CheckInitialization := FSetupValid
    AND FEqualResult.IsInitialized
    AND FNotEqualResult.IsInitialized
    AND FCaptureIntegrity.IsInitialized
    AND FFindingDetails.IsInitialized;
IF NOT CheckInitialization THEN
    EventPublisher.PublishEvent(Event := CreateFrameworkEvent(Name := Name,
        ResourceName := '',
        State := State,
        Severity := E_EventSeverity.Error,
        Message := 'Tolerance selftest setup failed.'));
END_IF;
END_METHOD

{region 'Documentation'}
(*!
<summary>Checks literal results, finding count and isolated finding identities.</summary>
*)
{endregion}
METHOD PRIVATE CheckResults
VAR
    FindingIndex : UINT;
    NotEqualFindingMatches : BOOL;
END_VAR
FEqualResultMatches := FEqualSubject.Result = FExpectedEqualResult;
FNotEqualResultMatches := FNotEqualSubject.Result = FExpectedNotEqualResult;
FCaptureIntegrityMatches := (FCaptureStatus.SequenceId = FExpectedFindings)
    AND (FCaptureStatus.LostEventCount = 0);

FindingIndex := 1;
FFindingDetailsMatch := TRUE;
IF FExpectedEqualFinding <> E_Result.NotEvaluated THEN
    FFindingDetailsMatch := IsFindingValid(Index := FindingIndex,
        ExpectedName := FEqualSubject.Name,
        ExpectedResult := FExpectedEqualFinding);
    FindingIndex := FindingIndex + 1;
END_IF;
IF FExpectedNotEqualFinding <> E_Result.NotEvaluated THEN
    NotEqualFindingMatches := IsFindingValid(Index := FindingIndex,
        ExpectedName := FNotEqualSubject.Name,
        ExpectedResult := FExpectedNotEqualFinding);
    FFindingDetailsMatch := FFindingDetailsMatch AND NotEqualFindingMatches;
END_IF;
END_METHOD

{region 'Documentation'}
(*!
<summary>Configures checking Assertions; subject actions remain in the test script.</summary>
*)
{endregion}
METHOD PROTECTED Configure
VAR
    Initialized : BOOL;
END_VAR
FPreparationStateCount := 0;
FTestStateCount := 1;
FEqualResult.Initialize(Parent := THIS^,
    AssertionName := 'EqualResult');
FNotEqualResult.Initialize(Parent := THIS^,
    AssertionName := 'NotEqualResult');
FCaptureIntegrity.Initialize(Parent := THIS^,
    AssertionName := 'CaptureIntegrity');
FFindingDetails.Initialize(Parent := THIS^,
    AssertionName := 'FindingDetails');
FSetupValid := FCapture.Initialize(Buffer := FEvents,
    FifoControl := FCaptureFifo,
    Status := FCaptureStatus);
FEqualSubject.BindPublisher(Publisher := FCapture);
Initialized := FEqualSubject.Initialize(Parent := THIS^,
    AssertionName := 'EqualSubject');
FSetupValid := FSetupValid AND Initialized;
FNotEqualSubject.BindPublisher(Publisher := FCapture);
Initialized := FNotEqualSubject.Initialize(Parent := THIS^,
    AssertionName := 'NotEqualSubject');
FSetupValid := FSetupValid AND Initialized;
END_METHOD

{region 'Documentation'}
(*!
<summary>Reads one of at most two captured findings; caller supplies index 1 or 2.</summary>
*)
{endregion}
METHOD PRIVATE IsFindingValid : BOOL //! TRUE when the selected captured finding satisfies the scenario metadata and diagnostic checks.
VAR_INPUT
    Index : UINT; //! One-based index in the retained isolated event capture.
    ExpectedName : STRING(GVL_Constants.NameLength); //! Independently authored Assertion name expected in the selected finding.
    ExpectedResult : E_Result; //! Independently authored finding result.
END_VAR
IsFindingValid := (FEvents[Index].SequenceId = UINT_TO_UDINT(Index))
    AND (FEvents[Index].Name = ExpectedName)
    AND (FEvents[Index].OwnerScope = E_OwnerScope.Assertion)
    AND (FEvents[Index].EventType = E_EventType.Result)
    AND (FEvents[Index].State = E_State.Running)
    AND (FEvents[Index].Result = ExpectedResult)
    AND (FEvents[Index].Message <> '');
END_METHOD

{region 'Documentation'}
(*!
<summary>Completes abort without asynchronous resources.</summary>
*)
{endregion}
METHOD PROTECTED ProcessAbort
VAR_INPUT
    Enable : BOOL; //! Phase permission supplied by the owning Test Case; FALSE does not authorize progression, while observation may continue.
END_VAR
IF Enable THEN
    CompleteAbort();
END_IF;
END_METHOD

{region 'Documentation'}
(*!
<summary>Latches checked observations before the next script step may proceed.</summary>
*)
{endregion}
METHOD PROTECTED ProcessAssertions
VAR_INPUT
    Enable : BOOL; //! Phase permission supplied by the owning Test Case; FALSE does not authorize progression, while observation may continue.
END_VAR
VAR
    Evaluate : BOOL;
END_VAR
Evaluate := Enable AND FObservationReady;
FEqualResult(Enable := Evaluate,
    State := State,
    IN := FEqualResultMatches);
FNotEqualResult(Enable := Evaluate,
    State := State,
    IN := FNotEqualResultMatches);
FCaptureIntegrity(Enable := Evaluate,
    State := State,
    IN := FCaptureIntegrityMatches);
FFindingDetails(Enable := Evaluate,
    State := State,
    IN := FFindingDetailsMatch);
IF Evaluate THEN
    FChecked := TRUE;
END_IF;
END_METHOD

{region 'Documentation'}
(*!
<summary>No Preparation phase is required.</summary>
*)
{endregion}
METHOD PROTECTED ProcessPreparations
VAR_INPUT
    // SA0033: Required hook; this test has no Preparation phase.
    {attribute 'analysis' := '-33'}
    Enable : BOOL; //! Phase permission supplied by the owning Test Case; FALSE does not authorize progression, while observation may continue.
END_VAR
END_METHOD

{region 'Documentation'}
(*!
<summary>Restarts the script and resets the checking Assertions.</summary>
*)
{endregion}
METHOD PROTECTED ProcessReset
FRow := EqualValues;
FRowPrepared := FALSE;
FChecked := FALSE;
FObservationReady := FALSE;
FEqualResult.Reset();
FEqualResultMatches := TRUE;
FNotEqualResult.Reset();
FNotEqualResultMatches := TRUE;
FCaptureIntegrity.Reset();
FCaptureIntegrityMatches := TRUE;
FFindingDetails.Reset();
FFindingDetailsMatch := TRUE;
CompleteReset();
END_METHOD

{region 'Documentation'}
(*!
<summary>Advances one bounded script step per active PLC cycle.</summary>
*)
{endregion}
METHOD PROTECTED ProcessTests
VAR_INPUT
    Enable : BOOL; //! Phase permission supplied by the owning Test Case; FALSE does not authorize progression, while observation may continue.
END_VAR
IF NOT Enable THEN
    RETURN;
END_IF;

IF FChecked THEN
    FChecked := FALSE;
    FObservationReady := FALSE;
    IF FRow = LastRow THEN
        CompleteTests();
        RETURN;
    END_IF;
    FRow := FRow + 1;
    FRowPrepared := FALSE;
END_IF;

IF NOT FRowPrepared THEN
    SelectRow();
    FCapture.Reset();
    IF NOT FPreserveResults THEN
        ResetSubjects();
    END_IF;
    CallSubjects(Enable := FALSE);
    FRowPrepared := TRUE;
ELSE
    CallSubjects(Enable := TRUE);
    CheckResults();
    FObservationReady := TRUE;
END_IF;
END_METHOD

{region 'Documentation'}
(*!
<summary>Requests fresh subject results before the next disabled call.</summary>
*)
{endregion}
METHOD PRIVATE ResetSubjects
FEqualSubject.Reset();
FNotEqualSubject.Reset();
END_METHOD

{region 'Documentation'}
(*!
<summary>Selects literal expectations; only named escalation rows retain preceding subject results.</summary>
*)
{endregion}
METHOD PRIVATE SelectRow
FPreserveResults := FALSE;
FExpected := REAL#8.0;
CASE FRow OF
    EqualValues:
        FActual := REAL#8.0;
        FTolerance := REAL#0.5;
        FExpectedEqualResult := E_Result.Passed;
        FExpectedNotEqualResult := E_Result.Failed;
        FExpectedFindings := 1;
        FExpectedEqualFinding := E_Result.NotEvaluated;
        FExpectedNotEqualFinding := E_Result.Failed;
    InsideLower:
        FActual := REAL#7.75;
        FTolerance := REAL#0.5;
        FExpectedEqualResult := E_Result.Passed;
        FExpectedNotEqualResult := E_Result.Failed;
        FExpectedFindings := 1;
        FExpectedEqualFinding := E_Result.NotEvaluated;
        FExpectedNotEqualFinding := E_Result.Failed;
    InsideUpper:
        FActual := REAL#8.25;
        FTolerance := REAL#0.5;
        FExpectedEqualResult := E_Result.Passed;
        FExpectedNotEqualResult := E_Result.Failed;
        FExpectedFindings := 1;
        FExpectedEqualFinding := E_Result.NotEvaluated;
        FExpectedNotEqualFinding := E_Result.Failed;
    AtLowerBoundary:
        FActual := REAL#7.5;
        FTolerance := REAL#0.5;
        FExpectedEqualResult := E_Result.Passed;
        FExpectedNotEqualResult := E_Result.Failed;
        FExpectedFindings := 1;
        FExpectedEqualFinding := E_Result.NotEvaluated;
        FExpectedNotEqualFinding := E_Result.Failed;
    AtUpperBoundary:
        FActual := REAL#8.5;
        FTolerance := REAL#0.5;
        FExpectedEqualResult := E_Result.Passed;
        FExpectedNotEqualResult := E_Result.Failed;
        FExpectedFindings := 1;
        FExpectedEqualFinding := E_Result.NotEvaluated;
        FExpectedNotEqualFinding := E_Result.Failed;
    OutsideLower:
        FActual := REAL#7.25;
        FTolerance := REAL#0.5;
        FExpectedEqualResult := E_Result.Failed;
        FExpectedNotEqualResult := E_Result.Passed;
        FExpectedFindings := 1;
        FExpectedEqualFinding := E_Result.Failed;
        FExpectedNotEqualFinding := E_Result.NotEvaluated;
    OutsideUpper:
        FActual := REAL#8.75;
        FTolerance := REAL#0.5;
        FExpectedEqualResult := E_Result.Failed;
        FExpectedNotEqualResult := E_Result.Passed;
        FExpectedFindings := 1;
        FExpectedEqualFinding := E_Result.Failed;
        FExpectedNotEqualFinding := E_Result.NotEvaluated;
    ZeroToleranceEqual:
        FActual := REAL#8.0;
        FTolerance := REAL#0.0;
        FExpectedEqualResult := E_Result.Passed;
        FExpectedNotEqualResult := E_Result.Failed;
        FExpectedFindings := 1;
        FExpectedEqualFinding := E_Result.NotEvaluated;
        FExpectedNotEqualFinding := E_Result.Failed;
    ZeroToleranceDifferent:
        FActual := REAL#8.25;
        FTolerance := REAL#0.0;
        FExpectedEqualResult := E_Result.Failed;
        FExpectedNotEqualResult := E_Result.Passed;
        FExpectedFindings := 1;
        FExpectedEqualFinding := E_Result.Failed;
        FExpectedNotEqualFinding := E_Result.NotEvaluated;
    NegativeTolerance:
        FActual := REAL#8.0;
        FTolerance := REAL#-0.5;
        FExpectedEqualResult := E_Result.Error;
        FExpectedNotEqualResult := E_Result.Error;
        FExpectedFindings := 2;
        FExpectedEqualFinding := E_Result.Error;
        FExpectedNotEqualFinding := E_Result.Error;
    EqualFailureBeforeError:
        FActual := REAL#9.0;
        FTolerance := REAL#0.5;
        FExpectedEqualResult := E_Result.Failed;
        FExpectedNotEqualResult := E_Result.Passed;
        FExpectedFindings := 1;
        FExpectedEqualFinding := E_Result.Failed;
        FExpectedNotEqualFinding := E_Result.NotEvaluated;
    ErrorAfterEqualFailure:
        FActual := REAL#9.0;
        FTolerance := REAL#-0.5;
        FExpectedEqualResult := E_Result.Error;
        FExpectedNotEqualResult := E_Result.Error;
        FExpectedFindings := 2;
        FExpectedEqualFinding := E_Result.Error;
        FExpectedNotEqualFinding := E_Result.Error;
        FPreserveResults := TRUE;
    RepeatedError:
        FActual := REAL#9.0;
        FTolerance := REAL#-0.5;
        FExpectedEqualResult := E_Result.Error;
        FExpectedNotEqualResult := E_Result.Error;
        FExpectedFindings := 0;
        FExpectedEqualFinding := E_Result.NotEvaluated;
        FExpectedNotEqualFinding := E_Result.NotEvaluated;
        FPreserveResults := TRUE;
    ValidInputsAfterError:
        FActual := REAL#8.0;
        FTolerance := REAL#0.5;
        FExpectedEqualResult := E_Result.Error;
        FExpectedNotEqualResult := E_Result.Error;
        FExpectedFindings := 0;
        FExpectedEqualFinding := E_Result.NotEvaluated;
        FExpectedNotEqualFinding := E_Result.NotEvaluated;
        FPreserveResults := TRUE;
    NotEqualFailureBeforeError:
        FActual := REAL#8.0;
        FTolerance := REAL#0.5;
        FExpectedEqualResult := E_Result.Passed;
        FExpectedNotEqualResult := E_Result.Failed;
        FExpectedFindings := 1;
        FExpectedEqualFinding := E_Result.NotEvaluated;
        FExpectedNotEqualFinding := E_Result.Failed;
    ErrorAfterNotEqualFailure:
        FActual := REAL#8.0;
        FTolerance := REAL#-0.5;
        FExpectedEqualResult := E_Result.Error;
        FExpectedNotEqualResult := E_Result.Error;
        FExpectedFindings := 2;
        FExpectedEqualFinding := E_Result.Error;
        FExpectedNotEqualFinding := E_Result.Error;
        FPreserveResults := TRUE;
    ResetRestoresEvaluation:
        FActual := REAL#8.0;
        FTolerance := REAL#0.5;
        FExpectedEqualResult := E_Result.Passed;
        FExpectedNotEqualResult := E_Result.Failed;
        FExpectedFindings := 1;
        FExpectedEqualFinding := E_Result.NotEvaluated;
        FExpectedNotEqualFinding := E_Result.Failed;
ELSE
    Error(Message := 'Unknown tolerance test row.');
END_CASE;
END_METHOD

END_FUNCTION_BLOCK

// ---- SelfTests/TestCases/TestSuite_AssertionFloatingPoint/Test_AssertionTolerance_LReal.TcPOU
{region 'Documentation'}
(*!
<summary>Checks LREAL absolute tolerance boundaries and Error escalation in both relations.</summary>
<description>
Named rows separate independent comparisons by a disabled reset call.
Only explicitly marked escalation rows retain the preceding subject result.
Outer Assertions latch every observation before advancing to the next row.
All finite comparison values are exact binary fractions; expected results are literal.
ErrorAfterEqualFailure and ErrorAfterNotEqualFailure exercise each held-Failed guard.
RepeatedError and ValidInputsAfterError require held Error without another finding.
Intentional findings remain in the local capture; no production algorithm is copied.
</description>
*)
{endregion}
FUNCTION_BLOCK Test_AssertionTolerance_LReal EXTENDS TestCaseBase
VAR
    FEqualSubject : AssertEqualTolerance_LReal;
    FNotEqualSubject : AssertNotEqualTolerance_LReal;
    FActual : LREAL;
    FExpected : LREAL;
    FTolerance : LREAL;
    FExpectedEqualResult : E_Result;
    FExpectedNotEqualResult : E_Result;
    FExpectedFindings : UDINT;
    FExpectedEqualFinding : E_Result;
    FExpectedNotEqualFinding : E_Result;
    FCapture : EventBuffer;
    FEvents : ARRAY[1..CaptureLength] OF ST_Event;
    FCaptureFifo : ST_FifoStatus;
    FCaptureStatus : ST_EventBufferStatus;
    FRow : UINT;
    FRowPrepared : BOOL;
    FPreserveResults : BOOL;
    FObservationReady : BOOL;
    FChecked : BOOL;
    FSetupValid : BOOL;
END_VAR
VAR
    FEqualResult : AssertTrue;
    FEqualResultMatches : BOOL;
    FNotEqualResult : AssertTrue;
    FNotEqualResultMatches : BOOL;
    FCaptureIntegrity : AssertTrue;
    FCaptureIntegrityMatches : BOOL;
    FFindingDetails : AssertTrue;
    FFindingDetailsMatch : BOOL;
END_VAR
VAR CONSTANT
    CaptureLength : UINT := 8;
    EqualValues : UINT := 1;
    InsideLower : UINT := 2;
    InsideUpper : UINT := 3;
    AtLowerBoundary : UINT := 4;
    AtUpperBoundary : UINT := 5;
    OutsideLower : UINT := 6;
    OutsideUpper : UINT := 7;
    ZeroToleranceEqual : UINT := 8;
    ZeroToleranceDifferent : UINT := 9;
    NegativeTolerance : UINT := 10;
    EqualFailureBeforeError : UINT := 11;
    ErrorAfterEqualFailure : UINT := 12;
    RepeatedError : UINT := 13;
    ValidInputsAfterError : UINT := 14;
    NotEqualFailureBeforeError : UINT := 15;
    ErrorAfterNotEqualFailure : UINT := 16;
    ResetRestoresEvaluation : UINT := 17;
    LastRow : UINT := ResetRestoresEvaluation;
END_VAR

SUPER^();

{region 'Documentation'}
(*!
<summary>Collects only outer checking Assertions, never intentional subject findings.</summary>
*)
{endregion}
METHOD PROTECTED AggregateResults
VAR_INPUT
    Aggregator : I_ResultAggregator; //! Borrowed result sink owned by the outer Test Case; add this test's checking Assertions without resetting or retaining the sink.
END_VAR
Aggregator.AddProvider(Provider := FEqualResult);
Aggregator.AddProvider(Provider := FNotEqualResult);
Aggregator.AddProvider(Provider := FCaptureIntegrity);
Aggregator.AddProvider(Provider := FFindingDetails);
END_METHOD

{region 'Documentation'}
(*!
<summary>Calls each inherited production Assertion once using the selected row.</summary>
*)
{endregion}
METHOD PRIVATE CallSubjects
VAR_INPUT
    Enable : BOOL; //! Observation-enable input forwarded to the controlled Assertion subjects for this call.
END_VAR
FEqualSubject(Enable := Enable,
    State := E_State.Running,
    IN := FActual,
    Expected := FExpected,
    Tolerance := FTolerance);
FNotEqualSubject(Enable := Enable,
    State := E_State.Running,
    IN := FActual,
    Expected := FExpected,
    Tolerance := FTolerance);
END_METHOD

{region 'Documentation'}
(*!
<summary>Extends base validation with subject and checking-Assertion setup.</summary>
*)
{endregion}
METHOD PROTECTED CheckInitialization : BOOL //! TRUE when the inherited initialization check and this concrete fixture check both accept the setup.
CheckInitialization := SUPER^.CheckInitialization();
IF NOT CheckInitialization THEN
    RETURN;
END_IF;

CheckInitialization := FSetupValid
    AND FEqualResult.IsInitialized
    AND FNotEqualResult.IsInitialized
    AND FCaptureIntegrity.IsInitialized
    AND FFindingDetails.IsInitialized;
IF NOT CheckInitialization THEN
    EventPublisher.PublishEvent(Event := CreateFrameworkEvent(Name := Name,
        ResourceName := '',
        State := State,
        Severity := E_EventSeverity.Error,
        Message := 'Tolerance selftest setup failed.'));
END_IF;
END_METHOD

{region 'Documentation'}
(*!
<summary>Checks literal results, finding count and isolated finding identities.</summary>
*)
{endregion}
METHOD PRIVATE CheckResults
VAR
    FindingIndex : UINT;
    NotEqualFindingMatches : BOOL;
END_VAR
FEqualResultMatches := FEqualSubject.Result = FExpectedEqualResult;
FNotEqualResultMatches := FNotEqualSubject.Result = FExpectedNotEqualResult;
FCaptureIntegrityMatches := (FCaptureStatus.SequenceId = FExpectedFindings)
    AND (FCaptureStatus.LostEventCount = 0);

FindingIndex := 1;
FFindingDetailsMatch := TRUE;
IF FExpectedEqualFinding <> E_Result.NotEvaluated THEN
    FFindingDetailsMatch := IsFindingValid(Index := FindingIndex,
        ExpectedName := FEqualSubject.Name,
        ExpectedResult := FExpectedEqualFinding);
    FindingIndex := FindingIndex + 1;
END_IF;
IF FExpectedNotEqualFinding <> E_Result.NotEvaluated THEN
    NotEqualFindingMatches := IsFindingValid(Index := FindingIndex,
        ExpectedName := FNotEqualSubject.Name,
        ExpectedResult := FExpectedNotEqualFinding);
    FFindingDetailsMatch := FFindingDetailsMatch AND NotEqualFindingMatches;
END_IF;
END_METHOD

{region 'Documentation'}
(*!
<summary>Configures checking Assertions; subject actions remain in the test script.</summary>
*)
{endregion}
METHOD PROTECTED Configure
VAR
    Initialized : BOOL;
END_VAR
FPreparationStateCount := 0;
FTestStateCount := 1;
FEqualResult.Initialize(Parent := THIS^,
    AssertionName := 'EqualResult');
FNotEqualResult.Initialize(Parent := THIS^,
    AssertionName := 'NotEqualResult');
FCaptureIntegrity.Initialize(Parent := THIS^,
    AssertionName := 'CaptureIntegrity');
FFindingDetails.Initialize(Parent := THIS^,
    AssertionName := 'FindingDetails');
FSetupValid := FCapture.Initialize(Buffer := FEvents,
    FifoControl := FCaptureFifo,
    Status := FCaptureStatus);
FEqualSubject.BindPublisher(Publisher := FCapture);
Initialized := FEqualSubject.Initialize(Parent := THIS^,
    AssertionName := 'EqualSubject');
FSetupValid := FSetupValid AND Initialized;
FNotEqualSubject.BindPublisher(Publisher := FCapture);
Initialized := FNotEqualSubject.Initialize(Parent := THIS^,
    AssertionName := 'NotEqualSubject');
FSetupValid := FSetupValid AND Initialized;
END_METHOD

{region 'Documentation'}
(*!
<summary>Reads one of at most two captured findings; caller supplies index 1 or 2.</summary>
*)
{endregion}
METHOD PRIVATE IsFindingValid : BOOL //! TRUE when the selected captured finding satisfies the scenario metadata and diagnostic checks.
VAR_INPUT
    Index : UINT; //! One-based index in the retained isolated event capture.
    ExpectedName : STRING(GVL_Constants.NameLength); //! Independently authored Assertion name expected in the selected finding.
    ExpectedResult : E_Result; //! Independently authored finding result.
END_VAR
IsFindingValid := (FEvents[Index].SequenceId = UINT_TO_UDINT(Index))
    AND (FEvents[Index].Name = ExpectedName)
    AND (FEvents[Index].OwnerScope = E_OwnerScope.Assertion)
    AND (FEvents[Index].EventType = E_EventType.Result)
    AND (FEvents[Index].State = E_State.Running)
    AND (FEvents[Index].Result = ExpectedResult)
    AND (FEvents[Index].Message <> '');
END_METHOD

{region 'Documentation'}
(*!
<summary>Completes abort without asynchronous resources.</summary>
*)
{endregion}
METHOD PROTECTED ProcessAbort
VAR_INPUT
    Enable : BOOL; //! Phase permission supplied by the owning Test Case; FALSE does not authorize progression, while observation may continue.
END_VAR
IF Enable THEN
    CompleteAbort();
END_IF;
END_METHOD

{region 'Documentation'}
(*!
<summary>Latches checked observations before the next script step may proceed.</summary>
*)
{endregion}
METHOD PROTECTED ProcessAssertions
VAR_INPUT
    Enable : BOOL; //! Phase permission supplied by the owning Test Case; FALSE does not authorize progression, while observation may continue.
END_VAR
VAR
    Evaluate : BOOL;
END_VAR
Evaluate := Enable AND FObservationReady;
FEqualResult(Enable := Evaluate,
    State := State,
    IN := FEqualResultMatches);
FNotEqualResult(Enable := Evaluate,
    State := State,
    IN := FNotEqualResultMatches);
FCaptureIntegrity(Enable := Evaluate,
    State := State,
    IN := FCaptureIntegrityMatches);
FFindingDetails(Enable := Evaluate,
    State := State,
    IN := FFindingDetailsMatch);
IF Evaluate THEN
    FChecked := TRUE;
END_IF;
END_METHOD

{region 'Documentation'}
(*!
<summary>No Preparation phase is required.</summary>
*)
{endregion}
METHOD PROTECTED ProcessPreparations
VAR_INPUT
    // SA0033: Required hook; this test has no Preparation phase.
    {attribute 'analysis' := '-33'}
    Enable : BOOL; //! Phase permission supplied by the owning Test Case; FALSE does not authorize progression, while observation may continue.
END_VAR
END_METHOD

{region 'Documentation'}
(*!
<summary>Restarts the script and resets the checking Assertions.</summary>
*)
{endregion}
METHOD PROTECTED ProcessReset
FRow := EqualValues;
FRowPrepared := FALSE;
FChecked := FALSE;
FObservationReady := FALSE;
FEqualResult.Reset();
FEqualResultMatches := TRUE;
FNotEqualResult.Reset();
FNotEqualResultMatches := TRUE;
FCaptureIntegrity.Reset();
FCaptureIntegrityMatches := TRUE;
FFindingDetails.Reset();
FFindingDetailsMatch := TRUE;
CompleteReset();
END_METHOD

{region 'Documentation'}
(*!
<summary>Advances one bounded script step per active PLC cycle.</summary>
*)
{endregion}
METHOD PROTECTED ProcessTests
VAR_INPUT
    Enable : BOOL; //! Phase permission supplied by the owning Test Case; FALSE does not authorize progression, while observation may continue.
END_VAR
IF NOT Enable THEN
    RETURN;
END_IF;

IF FChecked THEN
    FChecked := FALSE;
    FObservationReady := FALSE;
    IF FRow = LastRow THEN
        CompleteTests();
        RETURN;
    END_IF;
    FRow := FRow + 1;
    FRowPrepared := FALSE;
END_IF;

IF NOT FRowPrepared THEN
    SelectRow();
    FCapture.Reset();
    IF NOT FPreserveResults THEN
        ResetSubjects();
    END_IF;
    CallSubjects(Enable := FALSE);
    FRowPrepared := TRUE;
ELSE
    CallSubjects(Enable := TRUE);
    CheckResults();
    FObservationReady := TRUE;
END_IF;
END_METHOD

{region 'Documentation'}
(*!
<summary>Requests fresh subject results before the next disabled call.</summary>
*)
{endregion}
METHOD PRIVATE ResetSubjects
FEqualSubject.Reset();
FNotEqualSubject.Reset();
END_METHOD

{region 'Documentation'}
(*!
<summary>Selects literal expectations; only named escalation rows retain preceding subject results.</summary>
*)
{endregion}
METHOD PRIVATE SelectRow
FPreserveResults := FALSE;
FExpected := LREAL#8.0;
CASE FRow OF
    EqualValues:
        FActual := LREAL#8.0;
        FTolerance := LREAL#0.5;
        FExpectedEqualResult := E_Result.Passed;
        FExpectedNotEqualResult := E_Result.Failed;
        FExpectedFindings := 1;
        FExpectedEqualFinding := E_Result.NotEvaluated;
        FExpectedNotEqualFinding := E_Result.Failed;
    InsideLower:
        FActual := LREAL#7.75;
        FTolerance := LREAL#0.5;
        FExpectedEqualResult := E_Result.Passed;
        FExpectedNotEqualResult := E_Result.Failed;
        FExpectedFindings := 1;
        FExpectedEqualFinding := E_Result.NotEvaluated;
        FExpectedNotEqualFinding := E_Result.Failed;
    InsideUpper:
        FActual := LREAL#8.25;
        FTolerance := LREAL#0.5;
        FExpectedEqualResult := E_Result.Passed;
        FExpectedNotEqualResult := E_Result.Failed;
        FExpectedFindings := 1;
        FExpectedEqualFinding := E_Result.NotEvaluated;
        FExpectedNotEqualFinding := E_Result.Failed;
    AtLowerBoundary:
        FActual := LREAL#7.5;
        FTolerance := LREAL#0.5;
        FExpectedEqualResult := E_Result.Passed;
        FExpectedNotEqualResult := E_Result.Failed;
        FExpectedFindings := 1;
        FExpectedEqualFinding := E_Result.NotEvaluated;
        FExpectedNotEqualFinding := E_Result.Failed;
    AtUpperBoundary:
        FActual := LREAL#8.5;
        FTolerance := LREAL#0.5;
        FExpectedEqualResult := E_Result.Passed;
        FExpectedNotEqualResult := E_Result.Failed;
        FExpectedFindings := 1;
        FExpectedEqualFinding := E_Result.NotEvaluated;
        FExpectedNotEqualFinding := E_Result.Failed;
    OutsideLower:
        FActual := LREAL#7.25;
        FTolerance := LREAL#0.5;
        FExpectedEqualResult := E_Result.Failed;
        FExpectedNotEqualResult := E_Result.Passed;
        FExpectedFindings := 1;
        FExpectedEqualFinding := E_Result.Failed;
        FExpectedNotEqualFinding := E_Result.NotEvaluated;
    OutsideUpper:
        FActual := LREAL#8.75;
        FTolerance := LREAL#0.5;
        FExpectedEqualResult := E_Result.Failed;
        FExpectedNotEqualResult := E_Result.Passed;
        FExpectedFindings := 1;
        FExpectedEqualFinding := E_Result.Failed;
        FExpectedNotEqualFinding := E_Result.NotEvaluated;
    ZeroToleranceEqual:
        FActual := LREAL#8.0;
        FTolerance := LREAL#0.0;
        FExpectedEqualResult := E_Result.Passed;
        FExpectedNotEqualResult := E_Result.Failed;
        FExpectedFindings := 1;
        FExpectedEqualFinding := E_Result.NotEvaluated;
        FExpectedNotEqualFinding := E_Result.Failed;
    ZeroToleranceDifferent:
        FActual := LREAL#8.25;
        FTolerance := LREAL#0.0;
        FExpectedEqualResult := E_Result.Failed;
        FExpectedNotEqualResult := E_Result.Passed;
        FExpectedFindings := 1;
        FExpectedEqualFinding := E_Result.Failed;
        FExpectedNotEqualFinding := E_Result.NotEvaluated;
    NegativeTolerance:
        FActual := LREAL#8.0;
        FTolerance := LREAL#-0.5;
        FExpectedEqualResult := E_Result.Error;
        FExpectedNotEqualResult := E_Result.Error;
        FExpectedFindings := 2;
        FExpectedEqualFinding := E_Result.Error;
        FExpectedNotEqualFinding := E_Result.Error;
    EqualFailureBeforeError:
        FActual := LREAL#9.0;
        FTolerance := LREAL#0.5;
        FExpectedEqualResult := E_Result.Failed;
        FExpectedNotEqualResult := E_Result.Passed;
        FExpectedFindings := 1;
        FExpectedEqualFinding := E_Result.Failed;
        FExpectedNotEqualFinding := E_Result.NotEvaluated;
    ErrorAfterEqualFailure:
        FActual := LREAL#9.0;
        FTolerance := LREAL#-0.5;
        FExpectedEqualResult := E_Result.Error;
        FExpectedNotEqualResult := E_Result.Error;
        FExpectedFindings := 2;
        FExpectedEqualFinding := E_Result.Error;
        FExpectedNotEqualFinding := E_Result.Error;
        FPreserveResults := TRUE;
    RepeatedError:
        FActual := LREAL#9.0;
        FTolerance := LREAL#-0.5;
        FExpectedEqualResult := E_Result.Error;
        FExpectedNotEqualResult := E_Result.Error;
        FExpectedFindings := 0;
        FExpectedEqualFinding := E_Result.NotEvaluated;
        FExpectedNotEqualFinding := E_Result.NotEvaluated;
        FPreserveResults := TRUE;
    ValidInputsAfterError:
        FActual := LREAL#8.0;
        FTolerance := LREAL#0.5;
        FExpectedEqualResult := E_Result.Error;
        FExpectedNotEqualResult := E_Result.Error;
        FExpectedFindings := 0;
        FExpectedEqualFinding := E_Result.NotEvaluated;
        FExpectedNotEqualFinding := E_Result.NotEvaluated;
        FPreserveResults := TRUE;
    NotEqualFailureBeforeError:
        FActual := LREAL#8.0;
        FTolerance := LREAL#0.5;
        FExpectedEqualResult := E_Result.Passed;
        FExpectedNotEqualResult := E_Result.Failed;
        FExpectedFindings := 1;
        FExpectedEqualFinding := E_Result.NotEvaluated;
        FExpectedNotEqualFinding := E_Result.Failed;
    ErrorAfterNotEqualFailure:
        FActual := LREAL#8.0;
        FTolerance := LREAL#-0.5;
        FExpectedEqualResult := E_Result.Error;
        FExpectedNotEqualResult := E_Result.Error;
        FExpectedFindings := 2;
        FExpectedEqualFinding := E_Result.Error;
        FExpectedNotEqualFinding := E_Result.Error;
        FPreserveResults := TRUE;
    ResetRestoresEvaluation:
        FActual := LREAL#8.0;
        FTolerance := LREAL#0.5;
        FExpectedEqualResult := E_Result.Passed;
        FExpectedNotEqualResult := E_Result.Failed;
        FExpectedFindings := 1;
        FExpectedEqualFinding := E_Result.NotEvaluated;
        FExpectedNotEqualFinding := E_Result.Failed;
ELSE
    Error(Message := 'Unknown tolerance test row.');
END_CASE;
END_METHOD

END_FUNCTION_BLOCK

// ---- Framework/Assertions/POU/BasicTypes/LReal/AssertEqualTolerance_LReal.TcPOU
{region 'Documentation'}
(*!
<summary>Checks equality within absolute tolerance, including its boundary in
equality.</summary>
<description>

All checked operands and bounds must be finite; NaN or either infinity reports Error
during active evaluation.

Tolerance is absolute, in the same units as the values, finite and non-negative. Its
default zero requests exact comparison. The equality boundary is inclusive; larger differences
are unequal. Difference checking avoids overflow for large finite operands.

Numeric diagnostics use the formatter's default six significant digits; rounding affects
the message only, not the comparison.

</description>
*)
{endregion}
FUNCTION_BLOCK AssertEqualTolerance_LReal EXTENDS AssertionBase
VAR_INPUT
    IN : LREAL; //! Actual value checked or observed by this Assertion.
    Expected : LREAL; //! Reference value for comparison with IN.
    Tolerance : LREAL := 0.0; //! Maximum absolute difference accepted as equal; must be finite and non-negative.
END_VAR

SUPER^();

{region 'Documentation'}
(*!
<summary>Check equality within absolute tolerance, including its boundary in equality.</summary>
*)
{endregion}
METHOD PROTECTED Assert
VAR
    Message : STRING(GVL_Constants.MessageLength);
    ExpectedText : STRING(GVL_Constants.AssertionValueLength);
    ActualText : STRING(GVL_Constants.AssertionValueLength);
    ToleranceText : STRING(GVL_Constants.AssertionValueLength);
    IsWithinTolerance : BOOL;
END_VAR
IF NOT EvaluationActive THEN
    RETURN;
END_IF;

IF Result = E_Result.Error THEN
    RETURN;
END_IF;

IF NOT Tc2_Utilities.LrealIsFinite(x := IN) THEN
    Error(Message := 'Assertion error: IN must be finite.');
    RETURN;
END_IF;

IF NOT Tc2_Utilities.LrealIsFinite(x := Expected) THEN
    Error(Message := 'Assertion error: Expected must be finite.');
    RETURN;
END_IF;

IF NOT Tc2_Utilities.LrealIsFinite(x := Tolerance) THEN
    Error(Message := 'Assertion error: Tolerance must be finite.');
    RETURN;
END_IF;

IF Tolerance < 0.0 THEN
    ToleranceText := CreateAssertionTextValue_LReal(Value := Tolerance);
    Message := CONCAT('Assertion error: tolerance must not be negative. Tolerance = ',
        ToleranceText);
    Error(Message := Message);
    RETURN;
END_IF;

IF Result = E_Result.Failed THEN
    RETURN;
END_IF;

IsWithinTolerance := IsWithinTolerance_LReal(IN := IN,
    Expected := Expected,
    Tolerance := Tolerance);
IF NOT IsWithinTolerance THEN
    ExpectedText := CreateAssertionTextValue_LReal(Value := Expected);
    ActualText := CreateAssertionTextValue_LReal(Value := IN);
    ToleranceText := CreateAssertionTextValue_LReal(Value := Tolerance);
    Message := CONCAT('Assertion failed: values differ more than tolerance. Expected = ',
        ExpectedText);
    Message := CONCAT(Message, ', Actual = ');
    Message := CONCAT(Message, ActualText);
    Message := CONCAT(Message, ', Tolerance = ');
    Message := CONCAT(Message, ToleranceText);
    Message := CONCAT(Message, '.');
    Fail(Message := Message);
    RETURN;
END_IF;

Pass();
END_METHOD

END_FUNCTION_BLOCK

// ---- Framework/Assertions/POU/Utilities/CreateAssertionTextValue_LReal.TcPOU
{region 'Documentation'}
(*!
<summary>Formats LREAL diagnostics without floating-point arithmetic or native real-to-string conversion.</summary>
<description>Configurable significant decimal digits (default 6, clamped to 1..17), ties-to-even; NaN, +Inf, -Inf and signed zero are explicit.
Scientific notation keeps extreme values within AssertionValueLength. Does not determine Assertion validity.</description>
*)
{endregion}
FUNCTION INTERNAL CreateAssertionTextValue_LReal : STRING(GVL_Constants.AssertionValueLength) //! Bounded diagnostic text; not a value for subsequent numeric comparison.
VAR_INPUT
    Value : LREAL; //! Value to render as diagnostic text; formatting does not change comparison semantics.
    SignificantDigits : UINT := 6; //! Significant decimal digits; default 6, clamped to 1..17.
END_VAR
VAR
    Representation : AssertionLRealRepresentation;
    Fraction : ULINT;
    ExponentField : INT;
    Exponent : INT;
    Negative : BOOL;
END_VAR
VAR CONSTANT
    SignMask : LWORD := LWORD#16#8000000000000000;
    FractionMask : LWORD := LWORD#16#000FFFFFFFFFFFFF;
    ExponentMask : LWORD := LWORD#16#00000000000007FF;
    FractionBits : INT := 52;
    ExponentBias : INT := 1023;
    SpecialExponent : INT := 2047;
    ImplicitBit : ULINT := ULINT#4503599627370496;
    MaximumSignificantDigits : UINT := 17;
END_VAR

Representation.Value := Value;
Negative := (Representation.Bits AND SignMask) <> 0;
Fraction := LWORD_TO_ULINT(Representation.Bits AND FractionMask);
ExponentField := LWORD_TO_INT(SHR(Representation.Bits, FractionBits) AND ExponentMask);
IF ExponentField = SpecialExponent THEN
    IF Fraction <> 0 THEN
        CreateAssertionTextValue_LReal := 'NaN';
    ELSIF Negative THEN
        CreateAssertionTextValue_LReal := '-Inf';
    ELSE
        CreateAssertionTextValue_LReal := '+Inf';
    END_IF;
    RETURN;
END_IF;

IF ExponentField = 0 THEN
    Exponent := 1 - ExponentBias - FractionBits;
ELSE
    Fraction := Fraction + ImplicitBit;
    Exponent := ExponentField - ExponentBias - FractionBits;
END_IF;
CreateAssertionTextValue_LReal := CreateAssertionTextValue_BinaryFloat(Significand := Fraction,
    BinaryExponent := Exponent,
    Negative := Negative,
    SignificantDigits := UINT_TO_INT(LIMIT(UINT#1, SignificantDigits, MaximumSignificantDigits)));

END_FUNCTION

// ---- Framework/Assertions/POU/Utilities/CreateAssertionTextValue_BinaryFloat.TcPOU
{region 'Documentation'}
(*!
<summary>Formats an IEEE finite magnitude exactly before decimal rounding; used only by the typed diagnostic formatters.</summary>
<description>Preconditions: significand at most 53 bits; binary exponent -1074..971; precision 1..17.
Uses at most 86 base-1e9 limbs (344 bytes), 83 scale passes and bounded integer arithmetic.
No floating-point operation, dynamic allocation or full decimal expansion string.
Round-to-nearest, ties-to-even; trim fractional zeros and use scientific notation outside the compact fixed range.</description>
*)
{endregion}
FUNCTION INTERNAL CreateAssertionTextValue_BinaryFloat : STRING(GVL_Constants.AssertionValueLength) //! Bounded diagnostic text; not a value for subsequent numeric comparison.
VAR_INPUT
    Significand : ULINT; //! Unsigned binary significand, at most 53 bits; caller supplies a finite magnitude.
    BinaryExponent : INT; //! Power of two multiplying Significand; supported range -1074..971.
    Negative : BOOL; //! TRUE prefixes a minus sign, including negative zero.
    SignificantDigits : INT; //! Required significant decimal digits, 1..17; validated by the typed caller.
END_VAR
VAR
    Limbs : ARRAY[0..LimbCapacity - 1] OF UDINT;
    LimbCount : INT;
    LimbIndex : INT;
    RemainingExponent : INT;
    Scale : INT;
    Step : INT;
    StepLimit : INT;
    PowerBase : ULINT;
    Multiplier : ULINT;
    Carry : ULINT;
    Product : ULINT;
    LeadingDigits : ULINT;
    DigitCount : INT;
    TakenDigits : INT;
    DecimalExponent : INT;
    Divisor : ULINT;
    GuardDigit : ULINT;
    HasRemainder : BOOL;
    Digits : STRING(20);
    DigitLength : INT;
    DecimalPosition : INT;
    Text : STRING(GVL_Constants.AssertionValueLength);
    ExponentText : STRING(6);
    Index : INT;
END_VAR
VAR CONSTANT
    LimbCapacity : INT := 86;
    DecimalBase : ULINT := 1000000000;
    LimbDigits : INT := 9;
    BinaryChunk : INT := 29;
    FractionChunk : INT := 13;
    PowersOfTen : ARRAY[0..17] OF ULINT := [1, 10, 100, 1000, 10000, 100000, 1000000, 10000000, 100000000, 1000000000, 10000000000, 100000000000, 1000000000000, 10000000000000, 100000000000000, 1000000000000000, 10000000000000000, 100000000000000000];
END_VAR

IF Significand = 0 THEN
    IF Negative THEN
        CreateAssertionTextValue_BinaryFloat := '-0';
    ELSE
        CreateAssertionTextValue_BinaryFloat := '0';
    END_IF;
    RETURN;
END_IF;

{region 'Exact binary-to-decimal magnitude'}
Carry := Significand;
LimbCount := 0;
WHILE Carry <> 0 DO
    Limbs[LimbCount] := ULINT_TO_UDINT(Carry MOD DecimalBase);
    Carry := Carry / DecimalBase;
    LimbCount := LimbCount + 1;
END_WHILE;

Scale := 0;
PowerBase := 2;
StepLimit := BinaryChunk;
RemainingExponent := BinaryExponent;
IF BinaryExponent < 0 THEN
    // m * 2^-n = (m * 5^n) * 10^-n, including subnormal inputs.
    Scale := -BinaryExponent;
    PowerBase := 5;
    StepLimit := FractionChunk;
    RemainingExponent := Scale;
END_IF;

WHILE RemainingExponent > 0 DO
    Step := MIN(RemainingExponent, StepLimit);
    Multiplier := 1;
    FOR Index := 1 TO Step DO
        Multiplier := Multiplier * PowerBase;
    END_FOR;
    Carry := 0;
    FOR LimbIndex := 0 TO LimbCount - 1 DO
        Product := UDINT_TO_ULINT(Limbs[LimbIndex]) * Multiplier + Carry;
        Limbs[LimbIndex] := ULINT_TO_UDINT(Product MOD DecimalBase);
        Carry := Product / DecimalBase;
    END_FOR;
    WHILE Carry <> 0 DO
        Limbs[LimbCount] := ULINT_TO_UDINT(Carry MOD DecimalBase);
        Carry := Carry / DecimalBase;
        LimbCount := LimbCount + 1;
    END_WHILE;
    RemainingExponent := RemainingExponent - Step;
END_WHILE;
{endregion}

{region 'Significant digits and rounding'}
LimbIndex := LimbCount - 1;
LeadingDigits := UDINT_TO_ULINT(Limbs[LimbIndex]);
Digits := ULINT_TO_STRING(LeadingDigits);
DigitCount := LEN(Digits);
DecimalExponent := DigitCount + LimbDigits * LimbIndex - 1 - Scale;
HasRemainder := FALSE;
IF DigitCount > SignificantDigits + 1 THEN
    Divisor := PowersOfTen[DigitCount - SignificantDigits - 1];
    HasRemainder := (LeadingDigits MOD Divisor) <> 0;
    LeadingDigits := LeadingDigits / Divisor;
    DigitCount := SignificantDigits + 1;
END_IF;

WHILE (DigitCount < SignificantDigits + 1) AND (LimbIndex > 0) DO
    LimbIndex := LimbIndex - 1;
    TakenDigits := MIN(LimbDigits, SignificantDigits + 1 - DigitCount);
    Divisor := PowersOfTen[LimbDigits - TakenDigits];
    LeadingDigits := LeadingDigits * PowersOfTen[TakenDigits]
        + UDINT_TO_ULINT(Limbs[LimbIndex]) / Divisor;
    HasRemainder := (UDINT_TO_ULINT(Limbs[LimbIndex]) MOD Divisor) <> 0;
    DigitCount := DigitCount + TakenDigits;
END_WHILE;
FOR Index := 0 TO LimbIndex - 1 DO
    IF Limbs[Index] <> 0 THEN
        HasRemainder := TRUE;
        EXIT;
    END_IF;
END_FOR;

IF DigitCount > SignificantDigits THEN
    GuardDigit := LeadingDigits MOD 10;
    LeadingDigits := LeadingDigits / 10;
    IF (GuardDigit > 5)
        OR ((GuardDigit = 5) AND (HasRemainder OR ((LeadingDigits MOD 2) <> 0))) THEN
        LeadingDigits := LeadingDigits + 1;
    END_IF;
    IF LeadingDigits = PowersOfTen[SignificantDigits] THEN
        LeadingDigits := LeadingDigits / 10;
        DecimalExponent := DecimalExponent + 1;
    END_IF;
END_IF;

WHILE (LeadingDigits MOD 10) = 0 DO
    LeadingDigits := LeadingDigits / 10;
END_WHILE;
Digits := ULINT_TO_STRING(LeadingDigits);
DigitLength := LEN(Digits);
{endregion}

{region 'Bounded diagnostic text'}
IF (DecimalExponent >= 0) AND (DecimalExponent < SignificantDigits) THEN
    DecimalPosition := DecimalExponent + 1;
    IF DecimalPosition >= DigitLength THEN
        Text := Digits;
        FOR Index := DigitLength TO DecimalPosition - 1 DO
            Text := CONCAT(Text, '0');
        END_FOR;
    ELSE
        // SA0175: Generated ASCII decimal digits; split positions fit the current digit length.
        {analysis -175}
        Text := CONCAT(LEFT(Digits, DecimalPosition), '.');
        Text := CONCAT(Text, RIGHT(Digits, DigitLength - DecimalPosition));
        {analysis +175}
    END_IF;
ELSIF (DecimalExponent < 0) AND (DecimalExponent >= -4) THEN
    Text := '0.';
    FOR Index := 1 TO -DecimalExponent - 1 DO
        Text := CONCAT(Text, '0');
    END_FOR;
    Text := CONCAT(Text, Digits);
ELSE
    // SA0175: Generated ASCII decimal digits; split positions fit the current digit length.
    {analysis -175}
    Text := LEFT(Digits, 1);
    {analysis +175}
    IF DigitLength > 1 THEN
        Text := CONCAT(Text, '.');
        // SA0175: Generated ASCII decimal digits; split positions fit the current digit length.
        {analysis -175}
        Text := CONCAT(Text, RIGHT(Digits, DigitLength - 1));
        {analysis +175}
    END_IF;
    Text := CONCAT(Text, 'E');
    IF DecimalExponent >= 0 THEN
        Text := CONCAT(Text, '+');
    END_IF;
    ExponentText := INT_TO_STRING(DecimalExponent);
    Text := CONCAT(Text, ExponentText);
END_IF;
IF Negative THEN
    Text := CONCAT('-', Text);
END_IF;
CreateAssertionTextValue_BinaryFloat := Text;
{endregion}

END_FUNCTION

// ---- Framework/Assertions/POU/Utilities/IsWithinTolerance_LReal.TcPOU
{region 'Documentation'}
(*!
<summary>Tests absolute tolerance without overflowing the typed difference. Requires finite inputs and a finite, non-negative tolerance; the caller validates them.</summary>
*)
{endregion}
FUNCTION INTERNAL IsWithinTolerance_LReal : BOOL //! TRUE when the absolute difference is within Tolerance; caller must supply finite valid inputs.
VAR_INPUT
    IN : LREAL; //! Actual value checked or observed by this Assertion.
    Expected : LREAL; //! Reference value for comparison with IN.
    Tolerance : LREAL; //! Maximum absolute difference accepted as equal; must be finite and non-negative.
END_VAR
VAR
    ActualMagnitude : LREAL;
    ExpectedMagnitude : LREAL;
    LargeMagnitude : LREAL;
    SmallMagnitude : LREAL;
    RemainingMagnitude : LREAL;
    Difference : LREAL;
END_VAR
VAR CONSTANT
    MaxFinite : LREAL := LREAL#1.7976931348623157E308;
    HalfMaxFinite : LREAL := MaxFinite / LREAL#2.0;
END_VAR

IsWithinTolerance_LReal := FALSE;

IF ((IN < 0.0) AND (Expected > 0.0)) OR ((IN > 0.0) AND (Expected < 0.0)) THEN
    ActualMagnitude := ABS(IN);
    ExpectedMagnitude := ABS(Expected);
    LargeMagnitude := MAX(ActualMagnitude, ExpectedMagnitude);
    SmallMagnitude := MIN(ActualMagnitude, ExpectedMagnitude);

    IF LargeMagnitude >= HalfMaxFinite THEN
        // Exact subtraction: MaxFinite and LargeMagnitude are within a factor of two.
        RemainingMagnitude := MaxFinite - LargeMagnitude;
        IF SmallMagnitude > RemainingMagnitude THEN
            RETURN;
        END_IF;
    END_IF;
END_IF;

Difference := ABS(IN - Expected);
IsWithinTolerance_LReal := Difference <= Tolerance;

END_FUNCTION

// ---- Framework/Assertions/POU/BasicTypes/LReal/AssertNotEqualTolerance_LReal.TcPOU
{region 'Documentation'}
(*!
<summary>Checks inequality outside absolute tolerance, including its boundary in
equality.</summary>
<description>

All checked operands and bounds must be finite; NaN or either infinity reports Error
during active evaluation.

Tolerance is absolute, in the same units as the values, finite and non-negative. Its
default zero requests exact comparison. The equality boundary is inclusive; larger differences
are unequal. Difference checking avoids overflow for large finite operands.

Numeric diagnostics use the formatter's default six significant digits; rounding affects
the message only, not the comparison.

</description>
*)
{endregion}
FUNCTION_BLOCK AssertNotEqualTolerance_LReal EXTENDS AssertionBase
VAR_INPUT
    IN : LREAL; //! Actual value checked or observed by this Assertion.
    Expected : LREAL; //! Value that must differ from IN under this Assertion's comparison rules.
    Tolerance : LREAL := 0.0; //! Maximum absolute difference accepted as equal; must be finite and non-negative.
END_VAR

SUPER^();

{region 'Documentation'}
(*!
<summary>Check inequality outside absolute tolerance, including its boundary in equality.</summary>
*)
{endregion}
METHOD PROTECTED Assert
VAR
    Message : STRING(GVL_Constants.MessageLength);
    ExpectedText : STRING(GVL_Constants.AssertionValueLength);
    ActualText : STRING(GVL_Constants.AssertionValueLength);
    ToleranceText : STRING(GVL_Constants.AssertionValueLength);
    IsWithinTolerance : BOOL;
END_VAR
IF NOT EvaluationActive THEN
    RETURN;
END_IF;

IF Result = E_Result.Error THEN
    RETURN;
END_IF;

IF NOT Tc2_Utilities.LrealIsFinite(x := IN) THEN
    Error(Message := 'Assertion error: IN must be finite.');
    RETURN;
END_IF;

IF NOT Tc2_Utilities.LrealIsFinite(x := Expected) THEN
    Error(Message := 'Assertion error: Expected must be finite.');
    RETURN;
END_IF;

IF NOT Tc2_Utilities.LrealIsFinite(x := Tolerance) THEN
    Error(Message := 'Assertion error: Tolerance must be finite.');
    RETURN;
END_IF;

IF Tolerance < 0.0 THEN
    ToleranceText := CreateAssertionTextValue_LReal(Value := Tolerance);
    Message := CONCAT('Assertion error: tolerance must not be negative. Tolerance = ',
        ToleranceText);
    Error(Message := Message);
    RETURN;
END_IF;

IF Result = E_Result.Failed THEN
    RETURN;
END_IF;

IsWithinTolerance := IsWithinTolerance_LReal(IN := IN,
    Expected := Expected,
    Tolerance := Tolerance);
IF IsWithinTolerance THEN
    ExpectedText := CreateAssertionTextValue_LReal(Value := Expected);
    ActualText := CreateAssertionTextValue_LReal(Value := IN);
    ToleranceText := CreateAssertionTextValue_LReal(Value := Tolerance);
    Message := CONCAT('Assertion failed: values are equal within tolerance but should differ. NotExpected = ',
        ExpectedText);
    Message := CONCAT(Message, ', Actual = ');
    Message := CONCAT(Message, ActualText);
    Message := CONCAT(Message, ', Tolerance = ');
    Message := CONCAT(Message, ToleranceText);
    Message := CONCAT(Message, '.');
    Fail(Message := Message);
    RETURN;
END_IF;

Pass();
END_METHOD

END_FUNCTION_BLOCK

// ---- SelfTests/TestCases/TestSuite_AssertionFloatingPoint/Test_AssertionFiniteBoundaries_Real.TcPOU
{region 'Documentation'}
(*!
<summary>Checks REAL overflow-safe tolerance and representable precision boundaries.</summary>
<description>
Fixture representations are verified during configuration before any subject call.
MaxFinite versus -1 is mathematically outside every finite tolerance, even if rounded subtraction hides it.
The minimum-normal rows use zero or equal tolerance, without a denormal-mode assumption.
A disabled preparation call consumes subject resets before the next enabled observation.
Only outer checking Assertions contribute to the Test Case result.
Expected outcomes are explicit; production processing is inherited, not mirrored.
</description>
*)
{endregion}
FUNCTION_BLOCK Test_AssertionFiniteBoundaries_Real EXTENDS TestCaseBase
VAR
    FEqualSubject : AssertEqualTolerance_Real;
    FNotEqualSubject : AssertNotEqualTolerance_Real;
    FActual : REAL;
    FExpected : REAL;
    FTolerance : REAL;
    FMaximum : FloatingPointBits_Real;
    FHalfMaximum : FloatingPointBits_Real;
    FAdjacent : FloatingPointBits_Real;
    FGap : FloatingPointBits_Real;
    FHalfGap : FloatingPointBits_Real;
    FMinimumNormal : FloatingPointBits_Real;
    FExpectedEqualResult : E_Result;
    FExpectedNotEqualResult : E_Result;
    FExpectedFindings : UDINT;
    FCapture : EventBuffer;
    FEvents : ARRAY[1..CaptureLength] OF ST_Event;
    FCaptureFifo : ST_FifoStatus;
    FCaptureStatus : ST_EventBufferStatus;
    FRow : UINT;
    FRowPrepared : BOOL;
    FPreserveResults : BOOL;
    FObservationReady : BOOL;
    FChecked : BOOL;
    FSetupValid : BOOL;
END_VAR
VAR
    FEqualResult : AssertTrue;
    FEqualResultMatches : BOOL;
    FNotEqualResult : AssertTrue;
    FNotEqualResultMatches : BOOL;
    FCaptureIntegrity : AssertTrue;
    FCaptureIntegrityMatches : BOOL;
    FFindingDetails : AssertTrue;
    FFindingDetailsMatch : BOOL;
END_VAR
VAR CONSTANT
    CaptureLength : UINT := 8;
    FixtureSize : UINT := 4;
    OneBits : DWORD := DWORD#16#3F800000;
    MaximumBits : DWORD := DWORD#16#7F7FFFFF;
    HalfMaximumBits : DWORD := DWORD#16#7EFFFFFF;
    AdjacentBits : DWORD := DWORD#16#3F800001;
    GapBits : DWORD := DWORD#16#34000000;
    HalfGapBits : DWORD := DWORD#16#33800000;
    MinimumNormalBits : DWORD := DWORD#16#00800000;
    OppositeMaxima : UINT := 1;
    OppositeMaximaReversed : UINT := 2;
    MaximumAgainstZero : UINT := 3;
    MaximumAgainstNegativeOne : UINT := 4;
    NegativeOneAgainstMaximum : UINT := 5;
    EqualMaxima : UINT := 6;
    EqualNegativeMaxima : UINT := 7;
    OppositeBoundary : UINT := 8;
    BeyondOppositeBoundary : UINT := 9;
    LargeSameSignBoundary : UINT := 10;
    AdjacentAtTolerance : UINT := 11;
    AdjacentBelowTolerance : UINT := 12;
    AdjacentAtZero : UINT := 13;
    ReversedAdjacentBoundary : UINT := 14;
    MinimumNormalBoundary : UINT := 15;
    MinimumNormalAtZero : UINT := 16;
    NegativeMinimumNormal : UINT := 17;
    SmallOppositeBoundary : UINT := 18;
    SmallOppositeOutside : UINT := 19;
    LastRow : UINT := SmallOppositeOutside;
END_VAR

SUPER^();

{region 'Documentation'}
(*!
<summary>Collects only outer checking Assertions, never intentional subject findings.</summary>
*)
{endregion}
METHOD PROTECTED AggregateResults
VAR_INPUT
    Aggregator : I_ResultAggregator; //! Borrowed result sink owned by the outer Test Case; add this test's checking Assertions without resetting or retaining the sink.
END_VAR
Aggregator.AddProvider(Provider := FEqualResult);
Aggregator.AddProvider(Provider := FNotEqualResult);
Aggregator.AddProvider(Provider := FCaptureIntegrity);
Aggregator.AddProvider(Provider := FFindingDetails);
END_METHOD

{region 'Documentation'}
(*!
<summary>Calls each inherited production Assertion once using the selected row.</summary>
*)
{endregion}
METHOD PRIVATE CallSubjects
VAR_INPUT
    Enable : BOOL; //! Observation-enable input forwarded to the controlled Assertion subjects for this call.
END_VAR
FEqualSubject(Enable := Enable,
    State := E_State.Running,
    IN := FActual,
    Expected := FExpected,
    Tolerance := FTolerance);
FNotEqualSubject(Enable := Enable,
    State := E_State.Running,
    IN := FActual,
    Expected := FExpected,
    Tolerance := FTolerance);
END_METHOD

{region 'Documentation'}
(*!
<summary>Extends base validation with subject and checking-Assertion setup.</summary>
*)
{endregion}
METHOD PROTECTED CheckInitialization : BOOL //! TRUE when the inherited initialization check and this concrete fixture check both accept the setup.
CheckInitialization := SUPER^.CheckInitialization();
IF NOT CheckInitialization THEN
    RETURN;
END_IF;

CheckInitialization := FSetupValid
    AND FEqualResult.IsInitialized
    AND FNotEqualResult.IsInitialized
    AND FCaptureIntegrity.IsInitialized
    AND FFindingDetails.IsInitialized;
IF NOT CheckInitialization THEN
    EventPublisher.PublishEvent(Event := CreateFrameworkEvent(Name := Name,
        ResourceName := '',
        State := State,
        Severity := E_EventSeverity.Error,
        Message := 'Floating-point selftest setup or fixture representation failed.'));
END_IF;
END_METHOD

{region 'Documentation'}
(*!
<summary>Checks literal results and the ordered isolated findings from this row.</summary>
*)
{endregion}
METHOD PRIVATE CheckResults
VAR
    FindingIndex : UINT;
    FindingMatches : BOOL;
END_VAR
FEqualResultMatches := FEqualSubject.Result = FExpectedEqualResult;
FNotEqualResultMatches := FNotEqualSubject.Result = FExpectedNotEqualResult;
FCaptureIntegrityMatches := (FCaptureStatus.SequenceId = FExpectedFindings)
    AND (FCaptureStatus.LostEventCount = 0);

FindingIndex := 1;
FFindingDetailsMatch := TRUE;
IF (FExpectedEqualResult = E_Result.Failed) OR (FExpectedEqualResult = E_Result.Error) THEN
    FindingMatches := IsFindingValid(Index := FindingIndex,
        ExpectedName := FEqualSubject.Name,
        ExpectedResult := FExpectedEqualResult);
    FFindingDetailsMatch := FFindingDetailsMatch AND FindingMatches;
    FindingIndex := FindingIndex + 1;
END_IF;
IF (FExpectedNotEqualResult = E_Result.Failed) OR (FExpectedNotEqualResult = E_Result.Error) THEN
    FindingMatches := IsFindingValid(Index := FindingIndex,
        ExpectedName := FNotEqualSubject.Name,
        ExpectedResult := FExpectedNotEqualResult);
    FFindingDetailsMatch := FFindingDetailsMatch AND FindingMatches;
    FindingIndex := FindingIndex + 1;
END_IF;
END_METHOD

{region 'Documentation'}
(*!
<summary>Configures checking Assertions; subject actions remain in the test script.</summary>
*)
{endregion}
METHOD PROTECTED Configure
VAR
    Initialized : BOOL;
END_VAR
FPreparationStateCount := 0;
FTestStateCount := 1;
FSetupValid := InitializeValues();
FEqualResult.Initialize(Parent := THIS^,
    AssertionName := 'EqualResult');
FNotEqualResult.Initialize(Parent := THIS^,
    AssertionName := 'NotEqualResult');
FCaptureIntegrity.Initialize(Parent := THIS^,
    AssertionName := 'CaptureIntegrity');
FFindingDetails.Initialize(Parent := THIS^,
    AssertionName := 'FindingDetails');
Initialized := FCapture.Initialize(Buffer := FEvents,
    FifoControl := FCaptureFifo,
    Status := FCaptureStatus);
FSetupValid := FSetupValid AND Initialized;
FEqualSubject.BindPublisher(Publisher := FCapture);
Initialized := FEqualSubject.Initialize(Parent := THIS^,
    AssertionName := 'EqualSubject');
FSetupValid := FSetupValid AND Initialized;
FNotEqualSubject.BindPublisher(Publisher := FCapture);
Initialized := FNotEqualSubject.Initialize(Parent := THIS^,
    AssertionName := 'NotEqualSubject');
FSetupValid := FSetupValid AND Initialized;
END_METHOD

{region 'Documentation'}
(*!
<summary>Establishes typed fixtures and verifies their representation before any subject call.</summary>
*)
{endregion}
METHOD PRIVATE InitializeValues : BOOL //! TRUE when fixture sizes and floating-point bit representations match their explicit expected patterns.
VAR
    Representation : FloatingPointBits_Real;
END_VAR
Representation.Value := REAL#1.0;
InitializeValues := (SIZEOF(Representation) = FixtureSize)
    AND (Representation.Bits = OneBits);

FMaximum.Value := REAL#3.40282346638528859811704183484516925440E38;
Representation.Value := FMaximum.Value;
InitializeValues := InitializeValues AND (Representation.Bits = MaximumBits);
FHalfMaximum.Value := REAL#3.40282346638528859811704183484516925440E38 / REAL#2.0;
Representation.Value := FHalfMaximum.Value;
InitializeValues := InitializeValues AND (Representation.Bits = HalfMaximumBits);
FAdjacent.Value := REAL#1.00000011920928955078125;
Representation.Value := FAdjacent.Value;
InitializeValues := InitializeValues AND (Representation.Bits = AdjacentBits);
FGap.Value := REAL#1.1920928955078125E-7;
Representation.Value := FGap.Value;
InitializeValues := InitializeValues AND (Representation.Bits = GapBits);
FHalfGap.Value := REAL#1.1920928955078125E-7 / REAL#2.0;
Representation.Value := FHalfGap.Value;
InitializeValues := InitializeValues AND (Representation.Bits = HalfGapBits);
FMinimumNormal.Value := REAL#1.17549435082228750796873653722224568E-38;
Representation.Value := FMinimumNormal.Value;
InitializeValues := InitializeValues AND (Representation.Bits = MinimumNormalBits);
END_METHOD

{region 'Documentation'}
(*!
<summary>Reads a captured finding; the caller bounds the index by 2 subjects.</summary>
*)
{endregion}
METHOD PRIVATE IsFindingValid : BOOL //! TRUE when the selected captured finding satisfies the scenario metadata and diagnostic checks.
VAR_INPUT
    Index : UINT; //! One-based index in the retained isolated event capture.
    ExpectedName : STRING(GVL_Constants.NameLength); //! Independently authored Assertion name expected in the selected finding.
    ExpectedResult : E_Result; //! Independently authored finding result.
END_VAR
IsFindingValid := (FEvents[Index].SequenceId = UINT_TO_UDINT(Index))
    AND (FEvents[Index].Name = ExpectedName)
    AND (FEvents[Index].OwnerScope = E_OwnerScope.Assertion)
    AND (FEvents[Index].EventType = E_EventType.Result)
    AND (FEvents[Index].State = E_State.Running)
    AND (FEvents[Index].Result = ExpectedResult)
    AND (FEvents[Index].Message <> '');
END_METHOD

{region 'Documentation'}
(*!
<summary>Completes abort without asynchronous resources.</summary>
*)
{endregion}
METHOD PROTECTED ProcessAbort
VAR_INPUT
    Enable : BOOL; //! Phase permission supplied by the owning Test Case; FALSE does not authorize progression, while observation may continue.
END_VAR
IF Enable THEN
    CompleteAbort();
END_IF;
END_METHOD

{region 'Documentation'}
(*!
<summary>Latches checked observations before the next script step may proceed.</summary>
*)
{endregion}
METHOD PROTECTED ProcessAssertions
VAR_INPUT
    Enable : BOOL; //! Phase permission supplied by the owning Test Case; FALSE does not authorize progression, while observation may continue.
END_VAR
VAR
    Evaluate : BOOL;
END_VAR
Evaluate := Enable AND FObservationReady;
FEqualResult(Enable := Evaluate,
    State := State,
    IN := FEqualResultMatches);
FNotEqualResult(Enable := Evaluate,
    State := State,
    IN := FNotEqualResultMatches);
FCaptureIntegrity(Enable := Evaluate,
    State := State,
    IN := FCaptureIntegrityMatches);
FFindingDetails(Enable := Evaluate,
    State := State,
    IN := FFindingDetailsMatch);
IF Evaluate THEN
    FChecked := TRUE;
END_IF;
END_METHOD

{region 'Documentation'}
(*!
<summary>No Preparation phase is required.</summary>
*)
{endregion}
METHOD PROTECTED ProcessPreparations
VAR_INPUT
    // SA0033: Required hook; this test has no Preparation phase.
    {attribute 'analysis' := '-33'}
    Enable : BOOL; //! Phase permission supplied by the owning Test Case; FALSE does not authorize progression, while observation may continue.
END_VAR
END_METHOD

{region 'Documentation'}
(*!
<summary>Restarts the script and resets the checking Assertions.</summary>
*)
{endregion}
METHOD PROTECTED ProcessReset
FRow := OppositeMaxima;
FRowPrepared := FALSE;
FChecked := FALSE;
FObservationReady := FALSE;
FEqualResult.Reset();
FEqualResultMatches := TRUE;
FNotEqualResult.Reset();
FNotEqualResultMatches := TRUE;
FCaptureIntegrity.Reset();
FCaptureIntegrityMatches := TRUE;
FFindingDetails.Reset();
FFindingDetailsMatch := TRUE;
CompleteReset();
END_METHOD

{region 'Documentation'}
(*!
<summary>Advances one bounded script step per active PLC cycle.</summary>
*)
{endregion}
METHOD PROTECTED ProcessTests
VAR_INPUT
    Enable : BOOL; //! Phase permission supplied by the owning Test Case; FALSE does not authorize progression, while observation may continue.
END_VAR
IF NOT Enable THEN
    RETURN;
END_IF;

IF FChecked THEN
    FChecked := FALSE;
    FObservationReady := FALSE;
    IF FRow = LastRow THEN
        CompleteTests();
        RETURN;
    END_IF;
    FRow := FRow + 1;
    FRowPrepared := FALSE;
END_IF;

IF NOT FRowPrepared THEN
    SelectRow();
    FCapture.Reset();
    IF NOT FPreserveResults THEN
        ResetSubjects();
    END_IF;
    CallSubjects(Enable := FALSE);
    FRowPrepared := TRUE;
ELSE
    CallSubjects(Enable := TRUE);
    CheckResults();
    FObservationReady := TRUE;
END_IF;
END_METHOD

{region 'Documentation'}
(*!
<summary>Requests fresh subject results before the next disabled call.</summary>
*)
{endregion}
METHOD PRIVATE ResetSubjects
FEqualSubject.Reset();
FNotEqualSubject.Reset();
END_METHOD

{region 'Documentation'}
(*!
<summary>Selects independent literal outcomes; only named escalation rows preserve results.</summary>
*)
{endregion}
METHOD PRIVATE SelectRow
FPreserveResults := FALSE;
CASE FRow OF
    OppositeMaxima:
        FActual := FMaximum.Value;
        FExpected := -FMaximum.Value;
        FTolerance := FMaximum.Value;
        FExpectedEqualResult := E_Result.Failed;
        FExpectedNotEqualResult := E_Result.Passed;
        FExpectedFindings := 1;
    OppositeMaximaReversed:
        FActual := -FMaximum.Value;
        FExpected := FMaximum.Value;
        FTolerance := FMaximum.Value;
        FExpectedEqualResult := E_Result.Failed;
        FExpectedNotEqualResult := E_Result.Passed;
        FExpectedFindings := 1;
    MaximumAgainstZero:
        FActual := FMaximum.Value;
        FExpected := REAL#0.0;
        FTolerance := FMaximum.Value;
        FExpectedEqualResult := E_Result.Passed;
        FExpectedNotEqualResult := E_Result.Failed;
        FExpectedFindings := 1;
    MaximumAgainstNegativeOne:
        FActual := FMaximum.Value;
        FExpected := REAL#-1.0;
        FTolerance := FMaximum.Value;
        FExpectedEqualResult := E_Result.Failed;
        FExpectedNotEqualResult := E_Result.Passed;
        FExpectedFindings := 1;
    NegativeOneAgainstMaximum:
        FActual := REAL#-1.0;
        FExpected := FMaximum.Value;
        FTolerance := FMaximum.Value;
        FExpectedEqualResult := E_Result.Failed;
        FExpectedNotEqualResult := E_Result.Passed;
        FExpectedFindings := 1;
    EqualMaxima:
        FActual := FMaximum.Value;
        FExpected := FMaximum.Value;
        FTolerance := REAL#0.0;
        FExpectedEqualResult := E_Result.Passed;
        FExpectedNotEqualResult := E_Result.Failed;
        FExpectedFindings := 1;
    EqualNegativeMaxima:
        FActual := -FMaximum.Value;
        FExpected := -FMaximum.Value;
        FTolerance := REAL#0.0;
        FExpectedEqualResult := E_Result.Passed;
        FExpectedNotEqualResult := E_Result.Failed;
        FExpectedFindings := 1;
    OppositeBoundary:
        FActual := FHalfMaximum.Value;
        FExpected := -FHalfMaximum.Value;
        FTolerance := FMaximum.Value;
        FExpectedEqualResult := E_Result.Passed;
        FExpectedNotEqualResult := E_Result.Failed;
        FExpectedFindings := 1;
    BeyondOppositeBoundary:
        FActual := FHalfMaximum.Value;
        FExpected := -FMaximum.Value;
        FTolerance := FMaximum.Value;
        FExpectedEqualResult := E_Result.Failed;
        FExpectedNotEqualResult := E_Result.Passed;
        FExpectedFindings := 1;
    LargeSameSignBoundary:
        FActual := FMaximum.Value;
        FExpected := FHalfMaximum.Value;
        FTolerance := FHalfMaximum.Value;
        FExpectedEqualResult := E_Result.Passed;
        FExpectedNotEqualResult := E_Result.Failed;
        FExpectedFindings := 1;
    AdjacentAtTolerance:
        FActual := FAdjacent.Value;
        FExpected := REAL#1.0;
        FTolerance := FGap.Value;
        FExpectedEqualResult := E_Result.Passed;
        FExpectedNotEqualResult := E_Result.Failed;
        FExpectedFindings := 1;
    AdjacentBelowTolerance:
        FActual := FAdjacent.Value;
        FExpected := REAL#1.0;
        FTolerance := FHalfGap.Value;
        FExpectedEqualResult := E_Result.Failed;
        FExpectedNotEqualResult := E_Result.Passed;
        FExpectedFindings := 1;
    AdjacentAtZero:
        FActual := FAdjacent.Value;
        FExpected := REAL#1.0;
        FTolerance := REAL#0.0;
        FExpectedEqualResult := E_Result.Failed;
        FExpectedNotEqualResult := E_Result.Passed;
        FExpectedFindings := 1;
    ReversedAdjacentBoundary:
        FActual := REAL#1.0;
        FExpected := FAdjacent.Value;
        FTolerance := FGap.Value;
        FExpectedEqualResult := E_Result.Passed;
        FExpectedNotEqualResult := E_Result.Failed;
        FExpectedFindings := 1;
    MinimumNormalBoundary:
        FActual := FMinimumNormal.Value;
        FExpected := REAL#0.0;
        FTolerance := FMinimumNormal.Value;
        FExpectedEqualResult := E_Result.Passed;
        FExpectedNotEqualResult := E_Result.Failed;
        FExpectedFindings := 1;
    MinimumNormalAtZero:
        FActual := FMinimumNormal.Value;
        FExpected := REAL#0.0;
        FTolerance := REAL#0.0;
        FExpectedEqualResult := E_Result.Failed;
        FExpectedNotEqualResult := E_Result.Passed;
        FExpectedFindings := 1;
    NegativeMinimumNormal:
        FActual := -FMinimumNormal.Value;
        FExpected := REAL#0.0;
        FTolerance := FMinimumNormal.Value;
        FExpectedEqualResult := E_Result.Passed;
        FExpectedNotEqualResult := E_Result.Failed;
        FExpectedFindings := 1;
    SmallOppositeBoundary:
        FActual := REAL#1.0;
        FExpected := REAL#-1.0;
        FTolerance := REAL#2.0;
        FExpectedEqualResult := E_Result.Passed;
        FExpectedNotEqualResult := E_Result.Failed;
        FExpectedFindings := 1;
    SmallOppositeOutside:
        FActual := REAL#1.0;
        FExpected := REAL#-1.0;
        FTolerance := REAL#1.5;
        FExpectedEqualResult := E_Result.Failed;
        FExpectedNotEqualResult := E_Result.Passed;
        FExpectedFindings := 1;
ELSE
    Error(Message := 'Unknown floating-point test row.');
END_CASE;
END_METHOD

END_FUNCTION_BLOCK

// ---- SelfTests/TestCases/TestSuite_AssertionFloatingPoint/Test_AssertionFiniteBoundaries_LReal.TcPOU
{region 'Documentation'}
(*!
<summary>Checks LREAL overflow-safe tolerance and representable precision boundaries.</summary>
<description>
Fixture representations are verified during configuration before any subject call.
MaxFinite versus -1 is mathematically outside every finite tolerance, even if rounded subtraction hides it.
The minimum-normal rows use zero or equal tolerance, without a denormal-mode assumption.
A disabled preparation call consumes subject resets before the next enabled observation.
Only outer checking Assertions contribute to the Test Case result.
Expected outcomes are explicit; production processing is inherited, not mirrored.
</description>
*)
{endregion}
FUNCTION_BLOCK Test_AssertionFiniteBoundaries_LReal EXTENDS TestCaseBase
VAR
    FEqualSubject : AssertEqualTolerance_LReal;
    FNotEqualSubject : AssertNotEqualTolerance_LReal;
    FActual : LREAL;
    FExpected : LREAL;
    FTolerance : LREAL;
    FMaximum : FloatingPointBits_LReal;
    FHalfMaximum : FloatingPointBits_LReal;
    FAdjacent : FloatingPointBits_LReal;
    FGap : FloatingPointBits_LReal;
    FHalfGap : FloatingPointBits_LReal;
    FMinimumNormal : FloatingPointBits_LReal;
    FExpectedEqualResult : E_Result;
    FExpectedNotEqualResult : E_Result;
    FExpectedFindings : UDINT;
    FCapture : EventBuffer;
    FEvents : ARRAY[1..CaptureLength] OF ST_Event;
    FCaptureFifo : ST_FifoStatus;
    FCaptureStatus : ST_EventBufferStatus;
    FRow : UINT;
    FRowPrepared : BOOL;
    FPreserveResults : BOOL;
    FObservationReady : BOOL;
    FChecked : BOOL;
    FSetupValid : BOOL;
END_VAR
VAR
    FEqualResult : AssertTrue;
    FEqualResultMatches : BOOL;
    FNotEqualResult : AssertTrue;
    FNotEqualResultMatches : BOOL;
    FCaptureIntegrity : AssertTrue;
    FCaptureIntegrityMatches : BOOL;
    FFindingDetails : AssertTrue;
    FFindingDetailsMatch : BOOL;
END_VAR
VAR CONSTANT
    CaptureLength : UINT := 8;
    FixtureSize : UINT := 8;
    OneBits : LWORD := LWORD#16#3FF0000000000000;
    MaximumBits : LWORD := LWORD#16#7FEFFFFFFFFFFFFF;
    HalfMaximumBits : LWORD := LWORD#16#7FDFFFFFFFFFFFFF;
    AdjacentBits : LWORD := LWORD#16#3FF0000000000001;
    GapBits : LWORD := LWORD#16#3CB0000000000000;
    HalfGapBits : LWORD := LWORD#16#3CA0000000000000;
    MinimumNormalBits : LWORD := LWORD#16#0010000000000000;
    OppositeMaxima : UINT := 1;
    OppositeMaximaReversed : UINT := 2;
    MaximumAgainstZero : UINT := 3;
    MaximumAgainstNegativeOne : UINT := 4;
    NegativeOneAgainstMaximum : UINT := 5;
    EqualMaxima : UINT := 6;
    EqualNegativeMaxima : UINT := 7;
    OppositeBoundary : UINT := 8;
    BeyondOppositeBoundary : UINT := 9;
    LargeSameSignBoundary : UINT := 10;
    AdjacentAtTolerance : UINT := 11;
    AdjacentBelowTolerance : UINT := 12;
    AdjacentAtZero : UINT := 13;
    ReversedAdjacentBoundary : UINT := 14;
    MinimumNormalBoundary : UINT := 15;
    MinimumNormalAtZero : UINT := 16;
    NegativeMinimumNormal : UINT := 17;
    SmallOppositeBoundary : UINT := 18;
    SmallOppositeOutside : UINT := 19;
    LastRow : UINT := SmallOppositeOutside;
END_VAR

SUPER^();

{region 'Documentation'}
(*!
<summary>Collects only outer checking Assertions, never intentional subject findings.</summary>
*)
{endregion}
METHOD PROTECTED AggregateResults
VAR_INPUT
    Aggregator : I_ResultAggregator; //! Borrowed result sink owned by the outer Test Case; add this test's checking Assertions without resetting or retaining the sink.
END_VAR
Aggregator.AddProvider(Provider := FEqualResult);
Aggregator.AddProvider(Provider := FNotEqualResult);
Aggregator.AddProvider(Provider := FCaptureIntegrity);
Aggregator.AddProvider(Provider := FFindingDetails);
END_METHOD

{region 'Documentation'}
(*!
<summary>Calls each inherited production Assertion once using the selected row.</summary>
*)
{endregion}
METHOD PRIVATE CallSubjects
VAR_INPUT
    Enable : BOOL; //! Observation-enable input forwarded to the controlled Assertion subjects for this call.
END_VAR
FEqualSubject(Enable := Enable,
    State := E_State.Running,
    IN := FActual,
    Expected := FExpected,
    Tolerance := FTolerance);
FNotEqualSubject(Enable := Enable,
    State := E_State.Running,
    IN := FActual,
    Expected := FExpected,
    Tolerance := FTolerance);
END_METHOD

{region 'Documentation'}
(*!
<summary>Extends base validation with subject and checking-Assertion setup.</summary>
*)
{endregion}
METHOD PROTECTED CheckInitialization : BOOL //! TRUE when the inherited initialization check and this concrete fixture check both accept the setup.
CheckInitialization := SUPER^.CheckInitialization();
IF NOT CheckInitialization THEN
    RETURN;
END_IF;

CheckInitialization := FSetupValid
    AND FEqualResult.IsInitialized
    AND FNotEqualResult.IsInitialized
    AND FCaptureIntegrity.IsInitialized
    AND FFindingDetails.IsInitialized;
IF NOT CheckInitialization THEN
    EventPublisher.PublishEvent(Event := CreateFrameworkEvent(Name := Name,
        ResourceName := '',
        State := State,
        Severity := E_EventSeverity.Error,
        Message := 'Floating-point selftest setup or fixture representation failed.'));
END_IF;
END_METHOD

{region 'Documentation'}
(*!
<summary>Checks literal results and the ordered isolated findings from this row.</summary>
*)
{endregion}
METHOD PRIVATE CheckResults
VAR
    FindingIndex : UINT;
    FindingMatches : BOOL;
END_VAR
FEqualResultMatches := FEqualSubject.Result = FExpectedEqualResult;
FNotEqualResultMatches := FNotEqualSubject.Result = FExpectedNotEqualResult;
FCaptureIntegrityMatches := (FCaptureStatus.SequenceId = FExpectedFindings)
    AND (FCaptureStatus.LostEventCount = 0);

FindingIndex := 1;
FFindingDetailsMatch := TRUE;
IF (FExpectedEqualResult = E_Result.Failed) OR (FExpectedEqualResult = E_Result.Error) THEN
    FindingMatches := IsFindingValid(Index := FindingIndex,
        ExpectedName := FEqualSubject.Name,
        ExpectedResult := FExpectedEqualResult);
    FFindingDetailsMatch := FFindingDetailsMatch AND FindingMatches;
    FindingIndex := FindingIndex + 1;
END_IF;
IF (FExpectedNotEqualResult = E_Result.Failed) OR (FExpectedNotEqualResult = E_Result.Error) THEN
    FindingMatches := IsFindingValid(Index := FindingIndex,
        ExpectedName := FNotEqualSubject.Name,
        ExpectedResult := FExpectedNotEqualResult);
    FFindingDetailsMatch := FFindingDetailsMatch AND FindingMatches;
    FindingIndex := FindingIndex + 1;
END_IF;
END_METHOD

{region 'Documentation'}
(*!
<summary>Configures checking Assertions; subject actions remain in the test script.</summary>
*)
{endregion}
METHOD PROTECTED Configure
VAR
    Initialized : BOOL;
END_VAR
FPreparationStateCount := 0;
FTestStateCount := 1;
FSetupValid := InitializeValues();
FEqualResult.Initialize(Parent := THIS^,
    AssertionName := 'EqualResult');
FNotEqualResult.Initialize(Parent := THIS^,
    AssertionName := 'NotEqualResult');
FCaptureIntegrity.Initialize(Parent := THIS^,
    AssertionName := 'CaptureIntegrity');
FFindingDetails.Initialize(Parent := THIS^,
    AssertionName := 'FindingDetails');
Initialized := FCapture.Initialize(Buffer := FEvents,
    FifoControl := FCaptureFifo,
    Status := FCaptureStatus);
FSetupValid := FSetupValid AND Initialized;
FEqualSubject.BindPublisher(Publisher := FCapture);
Initialized := FEqualSubject.Initialize(Parent := THIS^,
    AssertionName := 'EqualSubject');
FSetupValid := FSetupValid AND Initialized;
FNotEqualSubject.BindPublisher(Publisher := FCapture);
Initialized := FNotEqualSubject.Initialize(Parent := THIS^,
    AssertionName := 'NotEqualSubject');
FSetupValid := FSetupValid AND Initialized;
END_METHOD

{region 'Documentation'}
(*!
<summary>Establishes typed fixtures and verifies their representation before any subject call.</summary>
*)
{endregion}
METHOD PRIVATE InitializeValues : BOOL //! TRUE when fixture sizes and floating-point bit representations match their explicit expected patterns.
VAR
    Representation : FloatingPointBits_LReal;
END_VAR
Representation.Value := LREAL#1.0;
InitializeValues := (SIZEOF(Representation) = FixtureSize)
    AND (Representation.Bits = OneBits);

FMaximum.Value := LREAL#1.7976931348623157E308;
Representation.Value := FMaximum.Value;
InitializeValues := InitializeValues AND (Representation.Bits = MaximumBits);
FHalfMaximum.Value := LREAL#1.7976931348623157E308 / LREAL#2.0;
Representation.Value := FHalfMaximum.Value;
InitializeValues := InitializeValues AND (Representation.Bits = HalfMaximumBits);
FAdjacent.Value := LREAL#1.0000000000000002220446049250313080847263336181640625;
Representation.Value := FAdjacent.Value;
InitializeValues := InitializeValues AND (Representation.Bits = AdjacentBits);
FGap.Value := LREAL#2.220446049250313080847263336181640625E-16;
Representation.Value := FGap.Value;
InitializeValues := InitializeValues AND (Representation.Bits = GapBits);
FHalfGap.Value := LREAL#2.220446049250313080847263336181640625E-16 / LREAL#2.0;
Representation.Value := FHalfGap.Value;
InitializeValues := InitializeValues AND (Representation.Bits = HalfGapBits);
FMinimumNormal.Value := LREAL#2.2250738585072014E-308;
Representation.Value := FMinimumNormal.Value;
InitializeValues := InitializeValues AND (Representation.Bits = MinimumNormalBits);
END_METHOD

{region 'Documentation'}
(*!
<summary>Reads a captured finding; the caller bounds the index by 2 subjects.</summary>
*)
{endregion}
METHOD PRIVATE IsFindingValid : BOOL //! TRUE when the selected captured finding satisfies the scenario metadata and diagnostic checks.
VAR_INPUT
    Index : UINT; //! One-based index in the retained isolated event capture.
    ExpectedName : STRING(GVL_Constants.NameLength); //! Independently authored Assertion name expected in the selected finding.
    ExpectedResult : E_Result; //! Independently authored finding result.
END_VAR
IsFindingValid := (FEvents[Index].SequenceId = UINT_TO_UDINT(Index))
    AND (FEvents[Index].Name = ExpectedName)
    AND (FEvents[Index].OwnerScope = E_OwnerScope.Assertion)
    AND (FEvents[Index].EventType = E_EventType.Result)
    AND (FEvents[Index].State = E_State.Running)
    AND (FEvents[Index].Result = ExpectedResult)
    AND (FEvents[Index].Message <> '');
END_METHOD

{region 'Documentation'}
(*!
<summary>Completes abort without asynchronous resources.</summary>
*)
{endregion}
METHOD PROTECTED ProcessAbort
VAR_INPUT
    Enable : BOOL; //! Phase permission supplied by the owning Test Case; FALSE does not authorize progression, while observation may continue.
END_VAR
IF Enable THEN
    CompleteAbort();
END_IF;
END_METHOD

{region 'Documentation'}
(*!
<summary>Latches checked observations before the next script step may proceed.</summary>
*)
{endregion}
METHOD PROTECTED ProcessAssertions
VAR_INPUT
    Enable : BOOL; //! Phase permission supplied by the owning Test Case; FALSE does not authorize progression, while observation may continue.
END_VAR
VAR
    Evaluate : BOOL;
END_VAR
Evaluate := Enable AND FObservationReady;
FEqualResult(Enable := Evaluate,
    State := State,
    IN := FEqualResultMatches);
FNotEqualResult(Enable := Evaluate,
    State := State,
    IN := FNotEqualResultMatches);
FCaptureIntegrity(Enable := Evaluate,
    State := State,
    IN := FCaptureIntegrityMatches);
FFindingDetails(Enable := Evaluate,
    State := State,
    IN := FFindingDetailsMatch);
IF Evaluate THEN
    FChecked := TRUE;
END_IF;
END_METHOD

{region 'Documentation'}
(*!
<summary>No Preparation phase is required.</summary>
*)
{endregion}
METHOD PROTECTED ProcessPreparations
VAR_INPUT
    // SA0033: Required hook; this test has no Preparation phase.
    {attribute 'analysis' := '-33'}
    Enable : BOOL; //! Phase permission supplied by the owning Test Case; FALSE does not authorize progression, while observation may continue.
END_VAR
END_METHOD

{region 'Documentation'}
(*!
<summary>Restarts the script and resets the checking Assertions.</summary>
*)
{endregion}
METHOD PROTECTED ProcessReset
FRow := OppositeMaxima;
FRowPrepared := FALSE;
FChecked := FALSE;
FObservationReady := FALSE;
FEqualResult.Reset();
FEqualResultMatches := TRUE;
FNotEqualResult.Reset();
FNotEqualResultMatches := TRUE;
FCaptureIntegrity.Reset();
FCaptureIntegrityMatches := TRUE;
FFindingDetails.Reset();
FFindingDetailsMatch := TRUE;
CompleteReset();
END_METHOD

{region 'Documentation'}
(*!
<summary>Advances one bounded script step per active PLC cycle.</summary>
*)
{endregion}
METHOD PROTECTED ProcessTests
VAR_INPUT
    Enable : BOOL; //! Phase permission supplied by the owning Test Case; FALSE does not authorize progression, while observation may continue.
END_VAR
IF NOT Enable THEN
    RETURN;
END_IF;

IF FChecked THEN
    FChecked := FALSE;
    FObservationReady := FALSE;
    IF FRow = LastRow THEN
        CompleteTests();
        RETURN;
    END_IF;
    FRow := FRow + 1;
    FRowPrepared := FALSE;
END_IF;

IF NOT FRowPrepared THEN
    SelectRow();
    FCapture.Reset();
    IF NOT FPreserveResults THEN
        ResetSubjects();
    END_IF;
    CallSubjects(Enable := FALSE);
    FRowPrepared := TRUE;
ELSE
    CallSubjects(Enable := TRUE);
    CheckResults();
    FObservationReady := TRUE;
END_IF;
END_METHOD

{region 'Documentation'}
(*!
<summary>Requests fresh subject results before the next disabled call.</summary>
*)
{endregion}
METHOD PRIVATE ResetSubjects
FEqualSubject.Reset();
FNotEqualSubject.Reset();
END_METHOD

{region 'Documentation'}
(*!
<summary>Selects independent literal outcomes; only named escalation rows preserve results.</summary>
*)
{endregion}
METHOD PRIVATE SelectRow
FPreserveResults := FALSE;
CASE FRow OF
    OppositeMaxima:
        FActual := FMaximum.Value;
        FExpected := -FMaximum.Value;
        FTolerance := FMaximum.Value;
        FExpectedEqualResult := E_Result.Failed;
        FExpectedNotEqualResult := E_Result.Passed;
        FExpectedFindings := 1;
    OppositeMaximaReversed:
        FActual := -FMaximum.Value;
        FExpected := FMaximum.Value;
        FTolerance := FMaximum.Value;
        FExpectedEqualResult := E_Result.Failed;
        FExpectedNotEqualResult := E_Result.Passed;
        FExpectedFindings := 1;
    MaximumAgainstZero:
        FActual := FMaximum.Value;
        FExpected := LREAL#0.0;
        FTolerance := FMaximum.Value;
        FExpectedEqualResult := E_Result.Passed;
        FExpectedNotEqualResult := E_Result.Failed;
        FExpectedFindings := 1;
    MaximumAgainstNegativeOne:
        FActual := FMaximum.Value;
        FExpected := LREAL#-1.0;
        FTolerance := FMaximum.Value;
        FExpectedEqualResult := E_Result.Failed;
        FExpectedNotEqualResult := E_Result.Passed;
        FExpectedFindings := 1;
    NegativeOneAgainstMaximum:
        FActual := LREAL#-1.0;
        FExpected := FMaximum.Value;
        FTolerance := FMaximum.Value;
        FExpectedEqualResult := E_Result.Failed;
        FExpectedNotEqualResult := E_Result.Passed;
        FExpectedFindings := 1;
    EqualMaxima:
        FActual := FMaximum.Value;
        FExpected := FMaximum.Value;
        FTolerance := LREAL#0.0;
        FExpectedEqualResult := E_Result.Passed;
        FExpectedNotEqualResult := E_Result.Failed;
        FExpectedFindings := 1;
    EqualNegativeMaxima:
        FActual := -FMaximum.Value;
        FExpected := -FMaximum.Value;
        FTolerance := LREAL#0.0;
        FExpectedEqualResult := E_Result.Passed;
        FExpectedNotEqualResult := E_Result.Failed;
        FExpectedFindings := 1;
    OppositeBoundary:
        FActual := FHalfMaximum.Value;
        FExpected := -FHalfMaximum.Value;
        FTolerance := FMaximum.Value;
        FExpectedEqualResult := E_Result.Passed;
        FExpectedNotEqualResult := E_Result.Failed;
        FExpectedFindings := 1;
    BeyondOppositeBoundary:
        FActual := FHalfMaximum.Value;
        FExpected := -FMaximum.Value;
        FTolerance := FMaximum.Value;
        FExpectedEqualResult := E_Result.Failed;
        FExpectedNotEqualResult := E_Result.Passed;
        FExpectedFindings := 1;
    LargeSameSignBoundary:
        FActual := FMaximum.Value;
        FExpected := FHalfMaximum.Value;
        FTolerance := FHalfMaximum.Value;
        FExpectedEqualResult := E_Result.Passed;
        FExpectedNotEqualResult := E_Result.Failed;
        FExpectedFindings := 1;
    AdjacentAtTolerance:
        FActual := FAdjacent.Value;
        FExpected := LREAL#1.0;
        FTolerance := FGap.Value;
        FExpectedEqualResult := E_Result.Passed;
        FExpectedNotEqualResult := E_Result.Failed;
        FExpectedFindings := 1;
    AdjacentBelowTolerance:
        FActual := FAdjacent.Value;
        FExpected := LREAL#1.0;
        FTolerance := FHalfGap.Value;
        FExpectedEqualResult := E_Result.Failed;
        FExpectedNotEqualResult := E_Result.Passed;
        FExpectedFindings := 1;
    AdjacentAtZero:
        FActual := FAdjacent.Value;
        FExpected := LREAL#1.0;
        FTolerance := LREAL#0.0;
        FExpectedEqualResult := E_Result.Failed;
        FExpectedNotEqualResult := E_Result.Passed;
        FExpectedFindings := 1;
    ReversedAdjacentBoundary:
        FActual := LREAL#1.0;
        FExpected := FAdjacent.Value;
        FTolerance := FGap.Value;
        FExpectedEqualResult := E_Result.Passed;
        FExpectedNotEqualResult := E_Result.Failed;
        FExpectedFindings := 1;
    MinimumNormalBoundary:
        FActual := FMinimumNormal.Value;
        FExpected := LREAL#0.0;
        FTolerance := FMinimumNormal.Value;
        FExpectedEqualResult := E_Result.Passed;
        FExpectedNotEqualResult := E_Result.Failed;
        FExpectedFindings := 1;
    MinimumNormalAtZero:
        FActual := FMinimumNormal.Value;
        FExpected := LREAL#0.0;
        FTolerance := LREAL#0.0;
        FExpectedEqualResult := E_Result.Failed;
        FExpectedNotEqualResult := E_Result.Passed;
        FExpectedFindings := 1;
    NegativeMinimumNormal:
        FActual := -FMinimumNormal.Value;
        FExpected := LREAL#0.0;
        FTolerance := FMinimumNormal.Value;
        FExpectedEqualResult := E_Result.Passed;
        FExpectedNotEqualResult := E_Result.Failed;
        FExpectedFindings := 1;
    SmallOppositeBoundary:
        FActual := LREAL#1.0;
        FExpected := LREAL#-1.0;
        FTolerance := LREAL#2.0;
        FExpectedEqualResult := E_Result.Passed;
        FExpectedNotEqualResult := E_Result.Failed;
        FExpectedFindings := 1;
    SmallOppositeOutside:
        FActual := LREAL#1.0;
        FExpected := LREAL#-1.0;
        FTolerance := LREAL#1.5;
        FExpectedEqualResult := E_Result.Failed;
        FExpectedNotEqualResult := E_Result.Passed;
        FExpectedFindings := 1;
ELSE
    Error(Message := 'Unknown floating-point test row.');
END_CASE;
END_METHOD

END_FUNCTION_BLOCK

// ---- SelfTests/TestCases/TestSuite_AssertionFloatingPoint/Test_AssertionRelations_Real.TcPOU
{region 'Documentation'}
(*!
<summary>Checks exact REAL ordering, inclusive ranges and signed zero.</summary>
<description>
Adjacent values differ by one representable step above 1; no implicit epsilon is allowed.
Range rows include both endpoints, equal bounds and invalid reversed bounds.
Extreme ordering uses comparisons only, not arithmetic differences.
A disabled preparation call consumes subject resets before the next enabled observation.
Only outer checking Assertions contribute to the Test Case result.
Expected outcomes are explicit; production processing is inherited, not mirrored.
</description>
*)
{endregion}
FUNCTION_BLOCK Test_AssertionRelations_Real EXTENDS TestCaseBase
VAR
    FEqualSubject : AssertEqual_Real;
    FNotEqualSubject : AssertNotEqual_Real;
    FLessThanSubject : AssertLessThan_Real;
    FLessEqualSubject : AssertLessEqual_Real;
    FGreaterThanSubject : AssertGreaterThan_Real;
    FGreaterEqualSubject : AssertGreaterEqual_Real;
    FInRangeSubject : AssertInRange_Real;
    FNotInRangeSubject : AssertNotInRange_Real;
    FActual : REAL;
    FExpected : REAL;
    FLower : REAL;
    FUpper : REAL;
    FMaximum : FloatingPointBits_Real;
    FAdjacent : FloatingPointBits_Real;
    FNegativeZero : FloatingPointBits_Real;
    FExpectedEqualResult : E_Result;
    FExpectedNotEqualResult : E_Result;
    FExpectedLessThanResult : E_Result;
    FExpectedLessEqualResult : E_Result;
    FExpectedGreaterThanResult : E_Result;
    FExpectedGreaterEqualResult : E_Result;
    FExpectedInRangeResult : E_Result;
    FExpectedNotInRangeResult : E_Result;
    FExpectedFindings : UDINT;
    FCapture : EventBuffer;
    FEvents : ARRAY[1..CaptureLength] OF ST_Event;
    FCaptureFifo : ST_FifoStatus;
    FCaptureStatus : ST_EventBufferStatus;
    FRow : UINT;
    FRowPrepared : BOOL;
    FPreserveResults : BOOL;
    FObservationReady : BOOL;
    FChecked : BOOL;
    FSetupValid : BOOL;
END_VAR
VAR
    FEqualResult : AssertTrue;
    FEqualResultMatches : BOOL;
    FNotEqualResult : AssertTrue;
    FNotEqualResultMatches : BOOL;
    FLessThanResult : AssertTrue;
    FLessThanResultMatches : BOOL;
    FLessEqualResult : AssertTrue;
    FLessEqualResultMatches : BOOL;
    FGreaterThanResult : AssertTrue;
    FGreaterThanResultMatches : BOOL;
    FGreaterEqualResult : AssertTrue;
    FGreaterEqualResultMatches : BOOL;
    FInRangeResult : AssertTrue;
    FInRangeResultMatches : BOOL;
    FNotInRangeResult : AssertTrue;
    FNotInRangeResultMatches : BOOL;
    FCaptureIntegrity : AssertTrue;
    FCaptureIntegrityMatches : BOOL;
    FFindingDetails : AssertTrue;
    FFindingDetailsMatch : BOOL;
END_VAR
VAR CONSTANT
    CaptureLength : UINT := 16;
    FixtureSize : UINT := 4;
    OneBits : DWORD := DWORD#16#3F800000;
    MaximumBits : DWORD := DWORD#16#7F7FFFFF;
    AdjacentBits : DWORD := DWORD#16#3F800001;
    NegativeZeroBits : DWORD := DWORD#16#80000000;
    EqualAtLowerBound : UINT := 1;
    AdjacentBelowExpected : UINT := 2;
    AdjacentAboveExpected : UINT := 3;
    Interior : UINT := 4;
    BelowRange : UINT := 5;
    AboveRange : UINT := 6;
    EqualBounds : UINT := 7;
    ReversedBounds : UINT := 8;
    SignedZero : UINT := 9;
    ExtremeAscending : UINT := 10;
    ExtremeDescending : UINT := 11;
    LastRow : UINT := ExtremeDescending;
END_VAR

SUPER^();

{region 'Documentation'}
(*!
<summary>Collects only outer checking Assertions, never intentional subject findings.</summary>
*)
{endregion}
METHOD PROTECTED AggregateResults
VAR_INPUT
    Aggregator : I_ResultAggregator; //! Borrowed result sink owned by the outer Test Case; add this test's checking Assertions without resetting or retaining the sink.
END_VAR
Aggregator.AddProvider(Provider := FEqualResult);
Aggregator.AddProvider(Provider := FNotEqualResult);
Aggregator.AddProvider(Provider := FLessThanResult);
Aggregator.AddProvider(Provider := FLessEqualResult);
Aggregator.AddProvider(Provider := FGreaterThanResult);
Aggregator.AddProvider(Provider := FGreaterEqualResult);
Aggregator.AddProvider(Provider := FInRangeResult);
Aggregator.AddProvider(Provider := FNotInRangeResult);
Aggregator.AddProvider(Provider := FCaptureIntegrity);
Aggregator.AddProvider(Provider := FFindingDetails);
END_METHOD

{region 'Documentation'}
(*!
<summary>Calls each inherited production Assertion once using the selected row.</summary>
*)
{endregion}
METHOD PRIVATE CallSubjects
VAR_INPUT
    Enable : BOOL; //! Observation-enable input forwarded to the controlled Assertion subjects for this call.
END_VAR
FEqualSubject(Enable := Enable,
    State := E_State.Running,
    IN := FActual,
    Expected := FExpected);
FNotEqualSubject(Enable := Enable,
    State := E_State.Running,
    IN := FActual,
    Expected := FExpected);
FLessThanSubject(Enable := Enable,
    State := E_State.Running,
    IN := FActual,
    Maximum := FExpected);
FLessEqualSubject(Enable := Enable,
    State := E_State.Running,
    IN := FActual,
    Maximum := FExpected);
FGreaterThanSubject(Enable := Enable,
    State := E_State.Running,
    IN := FActual,
    Minimum := FExpected);
FGreaterEqualSubject(Enable := Enable,
    State := E_State.Running,
    IN := FActual,
    Minimum := FExpected);
FInRangeSubject(Enable := Enable,
    State := E_State.Running,
    IN := FActual,
    Minimum := FLower,
    Maximum := FUpper);
FNotInRangeSubject(Enable := Enable,
    State := E_State.Running,
    IN := FActual,
    Minimum := FLower,
    Maximum := FUpper);
END_METHOD

{region 'Documentation'}
(*!
<summary>Extends base validation with subject and checking-Assertion setup.</summary>
*)
{endregion}
METHOD PROTECTED CheckInitialization : BOOL //! TRUE when the inherited initialization check and this concrete fixture check both accept the setup.
CheckInitialization := SUPER^.CheckInitialization();
IF NOT CheckInitialization THEN
    RETURN;
END_IF;

CheckInitialization := FSetupValid
    AND FEqualResult.IsInitialized
    AND FNotEqualResult.IsInitialized
    AND FLessThanResult.IsInitialized
    AND FLessEqualResult.IsInitialized
    AND FGreaterThanResult.IsInitialized
    AND FGreaterEqualResult.IsInitialized
    AND FInRangeResult.IsInitialized
    AND FNotInRangeResult.IsInitialized
    AND FCaptureIntegrity.IsInitialized
    AND FFindingDetails.IsInitialized;
IF NOT CheckInitialization THEN
    EventPublisher.PublishEvent(Event := CreateFrameworkEvent(Name := Name,
        ResourceName := '',
        State := State,
        Severity := E_EventSeverity.Error,
        Message := 'Floating-point selftest setup or fixture representation failed.'));
END_IF;
END_METHOD

{region 'Documentation'}
(*!
<summary>Checks literal results and the ordered isolated findings from this row.</summary>
*)
{endregion}
METHOD PRIVATE CheckResults
VAR
    FindingIndex : UINT;
    FindingMatches : BOOL;
END_VAR
FEqualResultMatches := FEqualSubject.Result = FExpectedEqualResult;
FNotEqualResultMatches := FNotEqualSubject.Result = FExpectedNotEqualResult;
FLessThanResultMatches := FLessThanSubject.Result = FExpectedLessThanResult;
FLessEqualResultMatches := FLessEqualSubject.Result = FExpectedLessEqualResult;
FGreaterThanResultMatches := FGreaterThanSubject.Result = FExpectedGreaterThanResult;
FGreaterEqualResultMatches := FGreaterEqualSubject.Result = FExpectedGreaterEqualResult;
FInRangeResultMatches := FInRangeSubject.Result = FExpectedInRangeResult;
FNotInRangeResultMatches := FNotInRangeSubject.Result = FExpectedNotInRangeResult;
FCaptureIntegrityMatches := (FCaptureStatus.SequenceId = FExpectedFindings)
    AND (FCaptureStatus.LostEventCount = 0);

FindingIndex := 1;
FFindingDetailsMatch := TRUE;
IF (FExpectedEqualResult = E_Result.Failed) OR (FExpectedEqualResult = E_Result.Error) THEN
    FindingMatches := IsFindingValid(Index := FindingIndex,
        ExpectedName := FEqualSubject.Name,
        ExpectedResult := FExpectedEqualResult);
    FFindingDetailsMatch := FFindingDetailsMatch AND FindingMatches;
    FindingIndex := FindingIndex + 1;
END_IF;
IF (FExpectedNotEqualResult = E_Result.Failed) OR (FExpectedNotEqualResult = E_Result.Error) THEN
    FindingMatches := IsFindingValid(Index := FindingIndex,
        ExpectedName := FNotEqualSubject.Name,
        ExpectedResult := FExpectedNotEqualResult);
    FFindingDetailsMatch := FFindingDetailsMatch AND FindingMatches;
    FindingIndex := FindingIndex + 1;
END_IF;
IF (FExpectedLessThanResult = E_Result.Failed) OR (FExpectedLessThanResult = E_Result.Error) THEN
    FindingMatches := IsFindingValid(Index := FindingIndex,
        ExpectedName := FLessThanSubject.Name,
        ExpectedResult := FExpectedLessThanResult);
    FFindingDetailsMatch := FFindingDetailsMatch AND FindingMatches;
    FindingIndex := FindingIndex + 1;
END_IF;
IF (FExpectedLessEqualResult = E_Result.Failed) OR (FExpectedLessEqualResult = E_Result.Error) THEN
    FindingMatches := IsFindingValid(Index := FindingIndex,
        ExpectedName := FLessEqualSubject.Name,
        ExpectedResult := FExpectedLessEqualResult);
    FFindingDetailsMatch := FFindingDetailsMatch AND FindingMatches;
    FindingIndex := FindingIndex + 1;
END_IF;
IF (FExpectedGreaterThanResult = E_Result.Failed) OR (FExpectedGreaterThanResult = E_Result.Error) THEN
    FindingMatches := IsFindingValid(Index := FindingIndex,
        ExpectedName := FGreaterThanSubject.Name,
        ExpectedResult := FExpectedGreaterThanResult);
    FFindingDetailsMatch := FFindingDetailsMatch AND FindingMatches;
    FindingIndex := FindingIndex + 1;
END_IF;
IF (FExpectedGreaterEqualResult = E_Result.Failed) OR (FExpectedGreaterEqualResult = E_Result.Error) THEN
    FindingMatches := IsFindingValid(Index := FindingIndex,
        ExpectedName := FGreaterEqualSubject.Name,
        ExpectedResult := FExpectedGreaterEqualResult);
    FFindingDetailsMatch := FFindingDetailsMatch AND FindingMatches;
    FindingIndex := FindingIndex + 1;
END_IF;
IF (FExpectedInRangeResult = E_Result.Failed) OR (FExpectedInRangeResult = E_Result.Error) THEN
    FindingMatches := IsFindingValid(Index := FindingIndex,
        ExpectedName := FInRangeSubject.Name,
        ExpectedResult := FExpectedInRangeResult);
    FFindingDetailsMatch := FFindingDetailsMatch AND FindingMatches;
    FindingIndex := FindingIndex + 1;
END_IF;
IF (FExpectedNotInRangeResult = E_Result.Failed) OR (FExpectedNotInRangeResult = E_Result.Error) THEN
    FindingMatches := IsFindingValid(Index := FindingIndex,
        ExpectedName := FNotInRangeSubject.Name,
        ExpectedResult := FExpectedNotInRangeResult);
    FFindingDetailsMatch := FFindingDetailsMatch AND FindingMatches;
    FindingIndex := FindingIndex + 1;
END_IF;
END_METHOD

{region 'Documentation'}
(*!
<summary>Configures checking Assertions; subject actions remain in the test script.</summary>
*)
{endregion}
METHOD PROTECTED Configure
VAR
    Initialized : BOOL;
END_VAR
FPreparationStateCount := 0;
FTestStateCount := 1;
FSetupValid := InitializeValues();
FEqualResult.Initialize(Parent := THIS^,
    AssertionName := 'EqualResult');
FNotEqualResult.Initialize(Parent := THIS^,
    AssertionName := 'NotEqualResult');
FLessThanResult.Initialize(Parent := THIS^,
    AssertionName := 'LessThanResult');
FLessEqualResult.Initialize(Parent := THIS^,
    AssertionName := 'LessEqualResult');
FGreaterThanResult.Initialize(Parent := THIS^,
    AssertionName := 'GreaterThanResult');
FGreaterEqualResult.Initialize(Parent := THIS^,
    AssertionName := 'GreaterEqualResult');
FInRangeResult.Initialize(Parent := THIS^,
    AssertionName := 'InRangeResult');
FNotInRangeResult.Initialize(Parent := THIS^,
    AssertionName := 'NotInRangeResult');
FCaptureIntegrity.Initialize(Parent := THIS^,
    AssertionName := 'CaptureIntegrity');
FFindingDetails.Initialize(Parent := THIS^,
    AssertionName := 'FindingDetails');
Initialized := FCapture.Initialize(Buffer := FEvents,
    FifoControl := FCaptureFifo,
    Status := FCaptureStatus);
FSetupValid := FSetupValid AND Initialized;
FEqualSubject.BindPublisher(Publisher := FCapture);
Initialized := FEqualSubject.Initialize(Parent := THIS^,
    AssertionName := 'EqualSubject');
FSetupValid := FSetupValid AND Initialized;
FNotEqualSubject.BindPublisher(Publisher := FCapture);
Initialized := FNotEqualSubject.Initialize(Parent := THIS^,
    AssertionName := 'NotEqualSubject');
FSetupValid := FSetupValid AND Initialized;
FLessThanSubject.BindPublisher(Publisher := FCapture);
Initialized := FLessThanSubject.Initialize(Parent := THIS^,
    AssertionName := 'LessThanSubject');
FSetupValid := FSetupValid AND Initialized;
FLessEqualSubject.BindPublisher(Publisher := FCapture);
Initialized := FLessEqualSubject.Initialize(Parent := THIS^,
    AssertionName := 'LessEqualSubject');
FSetupValid := FSetupValid AND Initialized;
FGreaterThanSubject.BindPublisher(Publisher := FCapture);
Initialized := FGreaterThanSubject.Initialize(Parent := THIS^,
    AssertionName := 'GreaterThanSubject');
FSetupValid := FSetupValid AND Initialized;
FGreaterEqualSubject.BindPublisher(Publisher := FCapture);
Initialized := FGreaterEqualSubject.Initialize(Parent := THIS^,
    AssertionName := 'GreaterEqualSubject');
FSetupValid := FSetupValid AND Initialized;
FInRangeSubject.BindPublisher(Publisher := FCapture);
Initialized := FInRangeSubject.Initialize(Parent := THIS^,
    AssertionName := 'InRangeSubject');
FSetupValid := FSetupValid AND Initialized;
FNotInRangeSubject.BindPublisher(Publisher := FCapture);
Initialized := FNotInRangeSubject.Initialize(Parent := THIS^,
    AssertionName := 'NotInRangeSubject');
FSetupValid := FSetupValid AND Initialized;
END_METHOD

{region 'Documentation'}
(*!
<summary>Establishes typed fixtures and verifies their representation before any subject call.</summary>
*)
{endregion}
METHOD PRIVATE InitializeValues : BOOL //! TRUE when fixture sizes and floating-point bit representations match their explicit expected patterns.
VAR
    Representation : FloatingPointBits_Real;
END_VAR
Representation.Value := REAL#1.0;
InitializeValues := (SIZEOF(Representation) = FixtureSize)
    AND (Representation.Bits = OneBits);

FMaximum.Value := REAL#3.40282346638528859811704183484516925440E38;
Representation.Value := FMaximum.Value;
InitializeValues := InitializeValues AND (Representation.Bits = MaximumBits);
FAdjacent.Value := REAL#1.00000011920928955078125;
Representation.Value := FAdjacent.Value;
InitializeValues := InitializeValues AND (Representation.Bits = AdjacentBits);
FNegativeZero.Bits := NegativeZeroBits;
Representation.Value := FNegativeZero.Value;
InitializeValues := InitializeValues AND (Representation.Bits = NegativeZeroBits);
END_METHOD

